(* IEC 61131-3 sources: daoli-st-library/DL_Device (part 7) *)

(* ---- I_DL_BarcodeScanner.st ---- *)
(*==============================================================================
 * 组件名称 (Component)  : I_DL_BarcodeScanner
 * 所属子库 (Sublibrary) : DL_Device
 * 当前版本 (Version)    : 1.0.0
 * 兼容性   (Platform)   : CODESYS 3.5 / TwinCAT 3 / 汇川 InoProShop / Machine Expert
 *                         纯 IEC 61131-3（第3版）接口语法，零厂商方言
 * 分类     (Category)   : 设备抽象接口（Interface）+ 配套状态枚举（DUT）
 * 功能简述 (Function)   : 工业固定式扫码枪标准抽象契约。路由分拣、批次追
 *                         溯、上下料校验等 DL_Process 模板的依赖注入件。
 *                         定义状态读取属性组（GET）与触发/应答/复位方法组；
 *                         串口/总线收发与数据本体由实现块（如
 *                         FB_DL_SerialScanner）经 IN_OUT 引脚注入，接口层
 *                         不做任何串口/总线收发与过程映像读写。
 * 契约结构 (Structure)  : 公约 0.11 接口三段式——状态枚举（本文件承载）+
 *                         属性（PROPERTY GET）+ 方法（METHOD）；方法共 3 个
 *                         （≤6 红线内）。故障态一律拒绝方法（红线：接口方
 *                         法拒绝语义），返回 FALSE 不静默成功。
 * 开源溯源 (Origin)     : 来源标签 tcopen-component / scanner-handshake
 *                         （RAW_NOTES_R7 S-2/S-3：TcOpen 组件接口分层思想
 *                         ——属性/方法分离契约与命令-应答握手语义，Apache
 *                         -2.0 公开资料，仅借鉴分层思想；接口命名、枚举编
 *                         号、方法签名 100% 本库独立设计，clean-room 未复
 *                         制源码）。
 * 归属说明 (Ownership)  : 本文件同时承载 E_DL_ScannerState 枚举定义，该枚
 *                         归属接口 I_DL_BarcodeScanner，与其同文件发布
 *                         （公约 0.11；禁止异文件同名异型重复定义）。
 * 红线自检 (Redline)    : R1 零全局变量表/外部变量引用 ✓｜R2 零物理 IO 地址 ✓
 *                         R3 纯 IEC 61131-3 ✓｜R4 N/A（契约件无运算）
 *                         R5 全成员中英双语同行注释 ✓｜R6 N/A（接口无状态机）
 *                         R7 N/A（无实例调用）｜R18 INTERFACE/END_INTERFACE
 *                         成对终结 ✓
 * 修订历史 (Revision)   :
 *   2026-11-15  v1.0.0  首版入库（Round 07 · DL_Device 扫码枪族接口件）
 *============================================================================*)

(*-----------------------------------------------------------------------------
 * 枚举: E_DL_ScannerState（归属接口 I_DL_BarcodeScanner，与其同文件）
 * 含义: 扫码枪握手状态机离散状态。编号步长 10 留空位便于后续插态而不破坏
 *       已有工程；eFault 取 99 保证排序末位（全库枚举编号惯例）。
 *----------------------------------------------------------------------------*)
TYPE E_DL_ScannerState :
(
    eIdle      := 0,    // 空闲待机：可受理解码触发 / Idle, ready to accept a decode trigger
    eTriggered := 10,   // 已触发：触发单拍输出已发出，等待下一拍进入读码 / Triggered, one-shot trigger output emitted
    eReading   := 20,   // 读码等待：结果窗口期内等待扫码枪回数 / Reading, waiting for the scanner reply inside the result window
    eOk        := 30,   // 解码成功：条码已锁存，等待应答消费 / Read OK, barcode latched, awaiting acknowledge
    eNoRead    := 40,   // 未读到：重试耗尽后的 NoRead 结果保持态 / NoRead, result hold state after retries exhausted
    eFault     := 99    // 故障锁存：连续 NoRead 超限/非法状态等，复位可尝试恢复 / Latched fault, reset may recover
) UINT;
END_TYPE

(*-----------------------------------------------------------------------------
 * 接口: I_DL_BarcodeScanner
 * 边界防错: 故障态一律拒绝方法；接口层不做任何串口/总线收发（数据本体经
 *           实现块 IN_OUT 引脚注入）；实现块负责握手编排与结果校验。
 *----------------------------------------------------------------------------*)
INTERFACE I_DL_BarcodeScanner

// ---- 属性段（全部只读 GET，实现块一一落地）----------------------------------

PROPERTY eState    : E_DL_ScannerState // 当前握手状态（Current handshake state），枚举见 E_DL_ScannerState
PROPERTY bReady    : BOOL              // 就绪可触发（Scanner ready），TRUE=处于可受理触发的状态 / TRUE = trigger acceptable
PROPERTY bReadOk   : BOOL              // 解码成功且结果有效（Read OK），TRUE=sBarcode 有效待消费 / TRUE = barcode valid and pending
PROPERTY bNoRead   : BOOL              // 未读到（NoRead），TRUE=重试耗尽未获得有效条码 / TRUE = no valid barcode after retries
PROPERTY sBarcode  : STRING(255)       // 最近有效条码字符串（Last valid barcode），长度 ≤255，bReadOk=TRUE 时有效 / Last valid barcode, valid when bReadOk
PROPERTY nReadCount: UDINT             // 累计成功解码次数（Total successful reads），复位不清零（追溯口径）/ Cumulative reads, preserved over reset
PROPERTY bFault    : BOOL              // 故障锁存中（Fault latched），显式排除信息级码（R21）/ TRUE = latched fault, info codes excluded
PROPERTY uErrorId  : UDINT             // 末次故障码（Last error code），0=无故障，段位 16#0003_xxxx / Last error code, family 16#0003_xxxx

// ---- 方法段（单发指令，返回受理/合法性结果）----------------------------------

METHOD CmdTrigger : BOOL // 触发一次解码（Trigger one decode），仅空闲态受理；非空闲/故障态拒绝返回 FALSE / Trigger one decode, accepted only in idle, rejected otherwise
VAR_INPUT
END_VAR

    END_METHOD

METHOD CmdAck : BOOL // 应答清除结果保持位（Acknowledge clears the result hold），eOk/eNoRead 态受理，为下一次解码前提 / Ack accepted in eOk/eNoRead
VAR_INPUT
END_VAR

    END_METHOD

METHOD CmdReset : BOOL // 复位故障（Reset fault），仅故障态受理返回 TRUE / Reset accepted only in fault state
VAR_INPUT
END_VAR

    END_METHOD
END_INTERFACE

(* ---- I_DL_Cylinder.st ---- *)
(*==============================================================================
 * 组件名称 (Component)  : I_DL_Cylinder
 * 所属子库 (Sublibrary) : DL_Device
 * 当前版本 (Version)    : 1.0.0
 * 兼容性   (Platform)   : CODESYS 3.5 / TwinCAT 3 / 汇川 InoProShop / Machine Expert
 *                         纯 IEC 61131-3（第3版）接口语法，零厂商方言
 * 分类     (Category)   : 设备抽象接口（Interface）+ 配套状态枚举（DUT）
 * 功能简述 (Function)   : 双电控气缸标准抽象契约。定义状态读取属性组（GET）与
 *                         动作指令方法组（Extend/Retract/Stop/Reset），供
 *                         DL_Process 全部机站动作层做依赖注入与解耦调用；
 *                         具体电磁阀输出与传感器采集由实现块（如
 *                         FB_DL_PneumaticCylinder）完成，接口层不做任何
 *                         过程映像读写，仅承载纯软件契约。
 * 开源溯源 (Origin)     : 来源标签 lbp-device（RAW_NOTES_R5 S-4：工业气动气缸
 *                         FB 设计指南 / LOGO! 气缸应用帖 / 双线圈互锁惯例，
 *                         公开教学文章，仅借鉴状态集合与故障分类等通用工程
 *                         语义；接口命名、方法签名按本库红线独立设计，
 *                         clean-room 未复制任何源码行）。
 * 红线自检 (Redline)    : R1 零全局变量表/外部变量引用 ✓｜R2 零物理 IO 地址 ✓
 *                         R3 纯 IEC 61131-3 ✓｜R5 全成员中英双语同行注释 ✓
 *                         R18 接口以 END_INTERFACE 成对终结 ✓
 * 归属说明 (Ownership)  : 本文件同时承载 E_DL_CylinderState 枚举定义，
 *                         该枚举归属接口 I_DL_Cylinder，与其同文件发布。
 * 修订历史 (Revision)   :
 *   2026-11-15  v1.0.0  首版入库（R5 轮 · DL_Device 开库）
 *============================================================================*)

(*-----------------------------------------------------------------------------
 * 枚举: E_DL_CylinderState（归属接口 I_DL_Cylinder，与其同文件）
 * 含义: 双电控气缸状态机离散状态。数值步长 10 留空位，便于后续插态
 *       而不破坏已有工程的持久化数值；eFault 取 99 保证排序末位。
 *----------------------------------------------------------------------------*)
TYPE E_DL_CylinderState :
(
    eIdle       := 0,    // 空闲稳态：双线圈全断，气缸保持当前位置 / Idle steady state, both coils off, cylinder holds position
    eExtending  := 10,   // 伸出动作中：伸出线圈得电，等待伸出到位反馈 / Extending, extend coil energized, waiting for extended feedback
    eExtended   := 20,   // 已伸出到位：伸出到位磁开确认的稳定终态 / Fully extended, confirmed by extended reed switch
    eRetracting := 30,   // 缩回动作中：缩回线圈得电，等待缩回到位反馈 / Retracting, retract coil energized, waiting for retracted feedback
    eRetracted  := 40,   // 已缩回到位：缩回到位磁开确认的稳定终态 / Fully retracted, confirmed by retracted reed switch
    eFault      := 99    // 故障锁存态：超时/传感器冲突/非法状态，仅复位可清 / Latched fault state, cleared only by reset
) UINT;
END_TYPE

(*-----------------------------------------------------------------------------
 * 接口: I_DL_Cylinder
 * 契约结构: 属性（PROPERTY GET）+ 方法（METHOD）两段式；方法总数 4 个，
 *           满足接口方法 ≤6 的拆分红线。所有方法均为非阻塞单发语义，
 *           不含跨扫描周期状态驻留；返回值仅表示"指令是否被受理"，
 *           实际动作完成以属性 eState/bExtended/bRetracted 为准。
 * 边界防错: 任何动作方法在故障锁存态一律拒绝并返回 FALSE；实现块负责
 *           信号采集与线圈驱动的全部过程映像交互，本接口不涉及。
 *----------------------------------------------------------------------------*)
INTERFACE I_DL_Cylinder

// ---- 属性段（全部只读 GET）------------------------------------------------

PROPERTY eState     : E_DL_CylinderState // 当前状态机状态（Current state）
PROPERTY bExtended  : BOOL               // 伸出到位磁开反馈（Extended reed feedback），TRUE=伸出到位
PROPERTY bRetracted : BOOL               // 缩回到位磁开反馈（Retracted reed feedback），TRUE=缩回到位
PROPERTY bFault     : BOOL               // 故障锁存中（Fault latched），TRUE=存在未复位故障
PROPERTY uErrorId   : UDINT              // 末次故障码（Last error code），0=无故障，段位 16#0003_xxxx

// ---- 方法段（单发指令，返回受理结果）--------------------------------------

METHOD CmdExtend : BOOL // 伸出指令（Extend command），单发；故障态拒绝返回 FALSE
VAR_INPUT
END_VAR

    END_METHOD

METHOD CmdRetract : BOOL // 缩回指令（Retract command），单发；故障态拒绝返回 FALSE
VAR_INPUT
END_VAR

    END_METHOD

METHOD CmdStop : BOOL // 停止指令（Stop command）：双线圈全断、保持当前位置；故障态拒绝返回 FALSE
VAR_INPUT
END_VAR

    END_METHOD

METHOD CmdReset : BOOL // 复位指令（Reset command），返回是否可复位（存在故障时为 TRUE）
VAR_INPUT
END_VAR

    END_METHOD
END_INTERFACE

(* ---- I_DL_FlowMeter.st ---- *)
(*==============================================================================
 * 组件名称 (Component)  : I_DL_FlowMeter
 * 所属子库 (Sublibrary) : DL_Device
 * 当前版本 (Version)    : 1.0.1
 * 兼容性   (Platform)   : CODESYS 3.5 / TwinCAT 3 / 汇川 InoProShop / Machine Expert
 *                         纯 IEC 61131-3（第3版）接口语法，零厂商方言
 * 分类     (Category)   : 设备抽象接口（Interface）+ 配套状态枚举（DUT）
 * 功能简述 (Function)   : 流量计标准抽象契约（脉冲型/模拟型均可适配）。定义
 *                         瞬时流量/累计总量读取属性组（GET）与总量清零/预置/
 *                         复位方法组，供批控与计量工站做依赖注入；脉冲采集
 *                         与频率估计由实现块（如 FB_DL_PulseFlowMeter）完成，
 *                         接口层不读物理输入。
 * 契约结构 (Structure)  : 公约 0.11 接口三段式——状态枚举（本文件承载）+
 *                         属性（PROPERTY GET）+ 方法（METHOD）；方法共 3 个
 *                         （≤6 红线内）。故障态一律拒绝方法。
 * 开源溯源 (Origin)     : 来源标签 tcopen-component / flow-totalizer
 *                         （RAW_NOTES_R7 S-2/S-6：TcOpen 组件接口分层思想与
 *                         工业流量计量公开语义域——瞬时流量/累计总量/低流
 *                         量截止，公开资料，仅借鉴语义域；接口命名、枚举编
 *                         号、方法签名 100% 本库独立设计，clean-room 未复
 *                         制源码）。
 * 归属说明 (Ownership)  : 本文件同时承载 E_DL_FlowMeterState 枚举定义，该枚
 *                         举归属接口 I_DL_FlowMeter，与其同文件发布（公约
 *                         0.11；禁止异文件同名异型重复定义）。
 * 红线自检 (Redline)    : R1 零全局变量表/外部变量引用 ✓｜R2 零物理 IO 地址 ✓
 *                         R3 纯 IEC 61131-3 ✓｜R4 N/A（契约件无运算）
 *                         R5 全成员中英双语同行注释 ✓｜R6 N/A（接口无状态机）
 *                         R7 N/A（无实例调用）｜R18 INTERFACE/END_INTERFACE
 *                         成对终结 ✓
 * 修订历史 (Revision)   :
 *   2026-11-15  v1.0.0  首版入库（Round 07 · DL_Device 流量计族接口件）
 *   2026-11-15  v1.0.1  R11 修复：枚举成员分隔符笔误，eFlowOk / eLowCutoff 两行误写单冒号 `:`（枚举成员赋值须用 `:=`），三平台编译阻断已消除，数值与语义不变。
 *                       R11 fix: enum member separator erratum, `:` -> `:=` on two members.
 *============================================================================*)

(*-----------------------------------------------------------------------------
 * 枚举: E_DL_FlowMeterState（归属接口 I_DL_FlowMeter，与其同文件）
 * 含义: 流量计量离散状态。编号步长 10 留空位，eFault 取 99 保证排序末位
 *       （全库枚举编号惯例）。
 *----------------------------------------------------------------------------*)
TYPE E_DL_FlowMeterState :
(
    eIdle      := 0,   // 空闲：未建窗或脉冲丢失超时后的静默态 / Idle, no window yet or silent after pulse timeout
    eMeasuring := 10,   // 测量中：采样窗运行中，流量待有效判定 / Measuring, sample window running, flow pending validation
    eFlowOk    := 20,  // 流量正常：高于低流量截止阈值的有效流量 / Flow OK, flow above the low-flow cutoff
    eLowCutoff := 30,  // 低流量截止：有效但低于阈值被截零（信息级）/ Low-flow cutoff, valid but zeroed below threshold (info)
    eFault     := 99   // 故障锁存：K 系数非法/非法状态，复位可尝试恢复 / Latched fault, reset may recover
) UINT;
END_TYPE

(*-----------------------------------------------------------------------------
 * 接口: I_DL_FlowMeter
 * 边界防错: 故障态一律拒绝方法并返回 FALSE；接口层不读物理输入；累计溢出
 *           防护（LREAL 整数精度边界预警）在实现块承载。
 *----------------------------------------------------------------------------*)
INTERFACE I_DL_FlowMeter

// ---- 属性段（全部只读 GET，实现块一一落地）----------------------------------

PROPERTY eState     : E_DL_FlowMeterState // 当前计量状态（Current metering state），枚举见 E_DL_FlowMeterState
PROPERTY fFlowRate  : REAL                // 瞬时流量（Flow rate）[L/min]，按 K 系数域换算 / Instantaneous flow rate [L/min], K-factor domain
PROPERTY fTotal     : LREAL               // 累计总量（Totalized volume）[L]，LREAL 防累计精度丢失 / Totalized volume [L], LREAL against precision loss
PROPERTY nPulseCount: UDINT               // 窗口内脉冲计数原始值（Pulse count of last window）/ Raw pulse count of the last window
PROPERTY bFault     : BOOL                // 故障锁存中（Fault latched），显式排除信息级码（R21）/ TRUE = latched fault, info codes excluded
PROPERTY uErrorId   : UDINT               // 末次故障码（Last error code），0=无故障，段位 16#0003_xxxx / Last error code, family 16#0003_xxxx

// ---- 方法段（单发指令，返回受理/合法性结果）----------------------------------

METHOD CmdTotalReset : BOOL // 总量清零（Total reset），批控切换零点；故障态拒绝 / Total reset, rejected in fault
VAR_INPUT
END_VAR

    END_METHOD

METHOD CmdTotalPreset : BOOL // 总量预置（Total preset），非有限值/负值拒绝 / Total preset, non-finite or negative rejected
VAR_INPUT
    fPreset : LREAL; // 预置总量（Preset volume）[L]，域 ≥0 / Preset volume [L], range >= 0
END_VAR

    END_METHOD

METHOD CmdReset : BOOL // 复位故障（Reset fault），仅故障态受理 / Reset accepted only in fault state
VAR_INPUT
END_VAR

    END_METHOD
END_INTERFACE

(* ---- I_DL_LevelSwitch.st ---- *)
(*==============================================================================
 * 组件名称 (Component)  : I_DL_LevelSwitch
 * 所属子库 (Sublibrary) : DL_Device
 * 当前版本 (Version)    : 1.0.0
 * 兼容性   (Platform)   : CODESYS 3.5 / TwinCAT 3 / 汇川 InoProShop / Machine Expert
 *                         纯 IEC 61131-3（第3版）接口语法，零厂商方言
 * 分类     (Category)   : 设备抽象接口（Interface）+ 配套状态枚举（DUT）
 * 功能简述 (Function)   : 料位开关标准抽象契约（振动叉/阻旋/电容等点式料位
 *                         开关通用）。高点溢流与低点干转联锁的统一契约；定
 *                         义有料判定/高/低联锁输出属性组（GET）与复位/测试
 *                         方法组；检测本体在传感器内部，接口层不做检测算法。
 * 契约结构 (Structure)  : 公约 0.11 接口三段式——状态枚举 + 失效安全模式枚
 *                         举（均本文件承载）+ 属性（PROPERTY GET）+ 方法
 *                         （METHOD）；方法共 2 个（≤6 红线内）。
 * 开源溯源 (Origin)     : 来源标签 tcopen-component / level-switch-failsafe
 *                         （RAW_NOTES_R7 S-2/S-7：TcOpen 组件接口分层思想与
 *                         料位开关失效安全公开语义域——fail-safe HIGH/LOW
 *                         方向约定、双联锁输出，公开资料，仅借鉴语义域；接
 *                         口命名、枚举编号、方法签名 100% 本库独立设计，
 *                         clean-room 未复制源码）。
 * 归属说明 (Ownership)  : 本文件同时承载 E_DL_LevelState 与 E_DL_FailSafeMode
 *                         两个枚举定义，均归属接口 I_DL_LevelSwitch，与其同
 *                         文件发布（公约 0.11；禁止异文件同名异型重复定义）。
 * 红线自检 (Redline)    : R1 零全局变量表/外部变量引用 ✓｜R2 零物理 IO 地址 ✓
 *                         R3 纯 IEC 61131-3 ✓｜R4 N/A（契约件无运算）
 *                         R5 全成员中英双语同行注释 ✓｜R6 N/A（接口无状态机）
 *                         R7 N/A（无实例调用）｜R18 INTERFACE/END_INTERFACE
 *                         成对终结 ✓
 * 修订历史 (Revision)   :
 *   2026-11-15  v1.0.0  首版入库（Round 07 · DL_Device 料位开关族接口件）
 *============================================================================*)

(*-----------------------------------------------------------------------------
 * 枚举: E_DL_LevelState（归属接口 I_DL_LevelSwitch，与其同文件）
 * 含义: 料位开关诊断状态。编号步长 10 留空位，eFault 取 99 保证排序末位
 *       （全库枚举编号惯例）。
 *----------------------------------------------------------------------------*)
TYPE E_DL_LevelState :
(
    eNoMaterial := 0,   // 无料：裸露确认态 / No material, bare confirmed
    eMaterial   := 10,  // 有料：覆盖确认态 / Material present, covered confirmed
    eSensorLoss := 20,  // 传感器失效态：按失效安全方向归一后的诊断镜像（本轮预留，检测算法后续轮次落地）/ Sensor loss, fail-safe normalized mirror (reserved this round)
    eFault      := 99   // 故障锁存：模式枚举越界等 / Latched fault
) UINT;
END_TYPE

(*-----------------------------------------------------------------------------
 * 枚举: E_DL_FailSafeMode（归属接口 I_DL_LevelSwitch，与其同文件）
 * 含义: 失效安全方向模式。决定传感器失效/使能切断时输出强制镜像的安全侧：
 *       eHigh=失效报有料（防溢流）；eLow=失效报无料（防干转）。
 *----------------------------------------------------------------------------*)
TYPE E_DL_FailSafeMode :
(
    eHigh := 0,   // 失效安全 HIGH：失效报有料，防溢流方向 / Fail-safe HIGH: failure reads covered, overflow protection
    eLow  := 1    // 失效安全 LOW：失效报无料，防干转方向 / Fail-safe LOW: failure reads bare, dry-run protection
) UINT;
END_TYPE

(*-----------------------------------------------------------------------------
 * 接口: I_DL_LevelSwitch
 * 边界防错: 故障态一律拒绝方法并返回 FALSE；接口层不做检测算法（检测本体
 *           在传感器内部）。
 *----------------------------------------------------------------------------*)
INTERFACE I_DL_LevelSwitch

// ---- 属性段（全部只读 GET，实现块一一落地）----------------------------------

PROPERTY eState    : E_DL_LevelState // 当前诊断状态（Current diagnostic state），枚举见 E_DL_LevelState
PROPERTY bMaterial : BOOL            // 有料判定输出（Material present），已按失效安全方向归一，TRUE=有料 / Fail-safe normalized material, TRUE = covered
PROPERTY bHighAlarm: BOOL            // 高点溢流联锁输出（High-level interlock），fail-safe HIGH 语义：归一有料即报警 / High alarm, fail-safe HIGH semantics
PROPERTY bLowAlarm : BOOL            // 低点干转联锁输出（Low-level interlock），fail-safe LOW 语义：归一无料即报警 / Low alarm, fail-safe LOW semantics
PROPERTY bFault    : BOOL            // 故障锁存中（Fault latched），显式排除信息级码（R21）/ TRUE = latched fault, info codes excluded
PROPERTY uErrorId  : UDINT           // 末次故障码（Last error code），0=无故障，段位 16#0003_xxxx / Last error code, family 16#0003_xxxx

// ---- 方法段（单发指令，返回受理/合法性结果）----------------------------------

METHOD CmdReset : BOOL // 复位故障（Reset fault），仅故障态受理 / Reset accepted only in fault state
VAR_INPUT
END_VAR

    END_METHOD

METHOD CmdTest : BOOL // 传感器功能测试请求（Sensor function test request），输出镜像进入测试态一拍 / Test request, test mirror asserted one scan
VAR_INPUT
END_VAR

    END_METHOD
END_INTERFACE

(* ---- I_DL_LightCurtain.st ---- *)
(*==============================================================================
 * 组件名称 (Component)  : I_DL_LightCurtain
 * 所属子库 (Sublibrary) : DL_Device
 * 当前版本 (Version)    : 1.0.0
 * 兼容性   (Platform)   : CODESYS 3.5 / TwinCAT 3 / 汇川 InoProShop / Machine Expert
 *                         纯 IEC 61131-3（第3版）接口语法，零厂商方言
 * 分类     (Category)   : 设备抽象接口（Interface）+ 配套状态枚举（DUT）
 * 功能简述 (Function)   : 安全光幕监控与屏蔽（Muting）标准抽象契约。定义光
 *                         幕状态读取属性组（GET）与滞留清除/确认/复位方法
 *                         组，供上层工站做依赖注入；OSSD 采集与屏蔽传感器
 *                         接线由实现块（如 FB_DL_SafetyLightCurtain）完成，
 *                         接口层不读物理输入。
 * 定位声明 (Positioning): 公约 0.13——本接口及其实现块为标准 PLC 逻辑编排
 *                         与诊断镜像层，不构成 ISO 13849 / IEC 62061 认证
 *                         安全功能，安全回路由认证安全控制器/安全 PLC 承载；
 *                         光幕本体 OSSD 的安全判断在认证安全光幕内部完成。
 * 契约结构 (Structure)  : 公约 0.11 接口三段式——状态枚举（本文件承载）+
 *                         属性（PROPERTY GET）+ 方法（METHOD）；方法共 3 个
 *                         （≤6 红线内）。故障态一律拒绝方法。
 * 边界防错 (Guard)      : bSafeStop 输出永不因屏蔽/override 置假——屏蔽态下
 *                         bSafeStop 断言恒 FALSE（光幕正常），实现块出口断
 *                         言承载。
 * 开源溯源 (Origin)     : 来源标签 tcopen-component / light-curtain-muting
 *                         （RAW_NOTES_R7 S-2/S-5：TcOpen 组件接口分层思想与
 *                         安全光幕屏蔽公开语义——OSSD 镜像、Muting/Override
 *                         状态域，公开资料，仅借鉴状态域语义；接口命名、枚
 *                         举编号、方法签名 100% 本库独立设计，clean-room 未
 *                         复制源码）。
 * 归属说明 (Ownership)  : 本文件同时承载 E_DL_CurtainState 枚举定义，该枚举
 *                         归属接口 I_DL_LightCurtain，与其同文件发布（公约
 *                         0.11；禁止异文件同名异型重复定义）。
 * 红线自检 (Redline)    : R1 零全局变量表/外部变量引用 ✓｜R2 零物理 IO 地址 ✓
 *                         R3 纯 IEC 61131-3 ✓｜R4 N/A（契约件无运算）
 *                         R5 全成员中英双语同行注释 ✓｜R6 N/A（接口无状态机）
 *                         R7 N/A（无实例调用）｜R18 INTERFACE/END_INTERFACE
 *                         成对终结 ✓
 * 修订历史 (Revision)   :
 *   2026-11-15  v1.0.0  首版入库（Round 07 · DL_Device 光幕族接口件）
 *============================================================================*)

(*-----------------------------------------------------------------------------
 * 枚举: E_DL_CurtainState（归属接口 I_DL_LightCurtain，与其同文件）
 * 含义: 光幕监控/屏蔽离散状态。编号步长 10 留空位，eFault 取 99 保证排序末
 *       位（全库枚举编号惯例）。
 *----------------------------------------------------------------------------*)
TYPE E_DL_CurtainState :
(
    eClear    := 0,   // 通光：光幕未被遮挡且无屏蔽活动 / Clear, curtain unblocked and no muting activity
    eBlocked  := 10,  // 遮挡：光幕被遮挡且未屏蔽（应停机镜像态）/ Blocked, curtain interrupted without muting (safe-stop mirror)
    eMuting   := 20,  // 屏蔽进行中：合法屏蔽序列屏蔽中 / Muting, a legal muting sequence is active
    eOverride := 30,   // 滞留清除进行中：钥匙开关滞留物清除 / Override, key-switch residual-object clearing active
    eFault    := 99   // 故障锁存：序列错误/屏蔽超时/OSSD 不一致/非法状态 / Latched fault
) UINT;
END_TYPE

(*-----------------------------------------------------------------------------
 * 接口: I_DL_LightCurtain
 * 边界防错: 故障态一律拒绝方法并返回 FALSE；bSafeStop 永不因屏蔽/override
 *           置假（屏蔽态下断言恒 FALSE，实现块承载）。
 *----------------------------------------------------------------------------*)
INTERFACE I_DL_LightCurtain

// ---- 属性段（全部只读 GET，实现块一一落地）----------------------------------

PROPERTY eState         : E_DL_CurtainState // 当前光幕状态（Current curtain state），枚举见 E_DL_CurtainState
PROPERTY bClear         : BOOL              // 光幕通光（Clear），OSSD 双通道全通光 / OSSD both channels clear
PROPERTY bMutingActive  : BOOL              // 屏蔽进行中（Muting active），合法屏蔽序列屏蔽中 / TRUE = legal muting sequence active
PROPERTY bOverrideActive: BOOL              // 滞留清除进行中（Override active），滞留物清除中 / TRUE = override clearing active
PROPERTY bSafeStop      : BOOL              // 应停机输出（Safe stop），光幕被遮挡且未屏蔽——本接口核心安全镜像位 / Curtain blocked and not muted, core safe-stop mirror
PROPERTY bFault         : BOOL              // 故障锁存中（Fault latched），显式排除信息级码（R21）/ TRUE = latched fault, info codes excluded
PROPERTY uErrorId       : UDINT             // 末次故障码（Last error code），0=无故障，段位 16#0003_xxxx / Last error code, family 16#0003_xxxx

// ---- 方法段（单发指令，返回受理/合法性结果）----------------------------------

METHOD CmdOverride : BOOL // 滞留物清除请求（Override request），前提至少一个屏蔽传感器仍遮挡，否则拒绝 / Override accepted only with at least one muting sensor blocked
VAR_INPUT
END_VAR

    END_METHOD

METHOD CmdAck : BOOL // 屏蔽/故障确认复位（Acknowledge of muting abort/fault），屏蔽序列中止后回评估态受理 / Ack after a muting abort, back to evaluation
VAR_INPUT
END_VAR

    END_METHOD

METHOD CmdReset : BOOL // 复位故障与重启联锁（Reset fault and restart interlock），仅故障态受理 / Reset accepted only in fault state
VAR_INPUT
END_VAR

    END_METHOD
END_INTERFACE

(* ---- I_DL_MotorDriver.st ---- *)
(*==============================================================================
 * 组件名称 (Component)  : I_DL_MotorDriver
 * 所属子库 (Sublibrary) : DL_Device
 * 当前版本 (Version)    : 1.0.0
 * 兼容性   (Platform)   : CODESYS 3.5 / TwinCAT 3 / 汇川 InoProShop / Machine Expert
 *                         纯 IEC 61131-3（第3版）接口语法，零厂商方言
 * 分类     (Category)   : 设备抽象接口（Interface）+ 配套状态枚举（DUT）
 * 功能简述 (Function)   : 直接启动（DOL）电机驱动器标准抽象契约。定义状态
 *                         读取属性组（GET，含重启抑制指示）与启停/复位方法组，
 *                         供机站动作层与配电监控层做依赖注入与解耦调用；
 *                         接触器线圈驱动与反馈采集由实现块（如 FB_DL_DolMotor）
 *                         完成，接口层不做任何过程映像读写。
 * 开源溯源 (Origin)     : 来源标签 lbp-device（RAW_NOTES_R5 S-4：DOL 电机保护
 *                         惯例——接触器反馈校验窗、热继电器过载锁存、防频繁
 *                         启停与重启抑制冷却时间为行业公知语义，公开教学
 *                         资料，仅借鉴通用工程语义；接口命名、方法签名按
 *                         本库红线独立设计，clean-room 未复制源码）。
 * 红线自检 (Redline)    : R1 零全局变量表/外部变量引用 ✓｜R2 零物理 IO 地址 ✓
 *                         R3 纯 IEC 61131-3 ✓｜R5 全成员中英双语同行注释 ✓
 *                         R18 接口以 END_INTERFACE 成对终结 ✓
 * 归属说明 (Ownership)  : 本文件同时承载 E_DL_MotorState 枚举定义，
 *                         该枚举归属接口 I_DL_MotorDriver，与其同文件发布。
 * 修订历史 (Revision)   :
 *   2026-11-15  v1.0.0  首版入库（R5 轮 · DL_Device 开库）
 *============================================================================*)

(*-----------------------------------------------------------------------------
 * 枚举: E_DL_MotorState（归属接口 I_DL_MotorDriver，与其同文件）
 * 含义: DOL 电机驱动状态机离散状态。数值步长 10 留空位，便于后续插态
 *       而不破坏已有工程的持久化数值；eFault 取 99 保证排序末位。
 *----------------------------------------------------------------------------*)
TYPE E_DL_MotorState :
(
    eIdle          := 0,    // 空闲停机态：接触器断开，可受理启动指令 / Idle stopped state, contactor open, start commands accepted
    eStarting      := 10,   // 启动校验态：线圈已得电，等待反馈窗内触点吸合确认 / Starting, coil energized, awaiting contactor pick-up confirmation within feedback window
    eRunning       := 20,   // 运行态：反馈吸合确认，正常带载运行 / Running, contactor feedback confirmed, loaded operation
    eStopping      := 30,   // 停机过渡态：线圈已断，等待反馈触点分断确认 / Stopping transition, coil de-energized, awaiting contactor drop-out confirmation
    eTripOverload  := 40,   // 过载脱扣态：热继电器动作锁存，仅复位且过载信号消失后可清 / Overload tripped and latched, cleared only by reset with overload signal removed
    eFault         := 99    // 故障锁存态：拒动/失反馈等故障，仅复位可清 / Latched fault state (refusal, feedback loss), cleared only by reset
) UINT;
END_TYPE

(*-----------------------------------------------------------------------------
 * 接口: I_DL_MotorDriver
 * 契约结构: 属性（PROPERTY GET）+ 方法（METHOD）两段式；方法总数 3 个，
 *           满足接口方法 ≤6 的拆分红线。所有方法均为非阻塞单发语义，
 *           不含跨扫描周期状态驻留；启动/复位方法返回值表示"指令是否
 *           被受理"，实际运行状态以属性 eState/bRunning 为准。
 * 边界防错: 启动方法在被抑制（重启抑制/次数超限）或故障态一律返回 FALSE；
 *           停止为无条件安全指令；实现块负责线圈驱动与触点反馈采集的
 *           全部过程映像交互，本接口不涉及。
 *----------------------------------------------------------------------------*)
INTERFACE I_DL_MotorDriver

// ---- 属性段（全部只读 GET）------------------------------------------------

PROPERTY eState          : E_DL_MotorState // 当前状态机状态（Current state）
PROPERTY bRunning        : BOOL            // 运行反馈（Running feedback），TRUE=反馈吸合确认运行中 / TRUE = running confirmed by contactor feedback
PROPERTY bFault          : BOOL            // 故障锁存中（Fault latched），TRUE=存在未复位故障（含过载脱扣）/ TRUE = latched fault incl. overload trip
PROPERTY uErrorId        : UDINT           // 末次故障码（Last error code），0=无故障，段位 16#0003_xxxx / Last error code, 0 = none, family 16#0003_xxxx
PROPERTY bRestartInhibit : BOOL            // 重启抑制激活中（Restart inhibit active），TRUE=冷却期内拒绝启动 / TRUE = start refused during cooling period

// ---- 方法段（单发指令，返回受理结果）--------------------------------------

METHOD CmdStart : BOOL // 启动指令（Start command），单发；被抑制/故障态返回 FALSE / Rejected with FALSE when inhibited or faulty
VAR_INPUT
END_VAR

    END_METHOD

METHOD CmdStop // 停止指令（Stop command），无条件安全动作，双线圈全断 / Unconditional safe stop command
VAR_INPUT
END_VAR

    END_METHOD

METHOD CmdReset : BOOL // 复位过载/故障（Reset overload and fault），返回是否可复位 / Returns TRUE only when resettable
VAR_INPUT
END_VAR

    END_METHOD
END_INTERFACE

(* ---- I_DL_MotorizedValve.st ---- *)
(*==============================================================================
 * 组件名称 (Component)  : I_DL_MotorizedValve
 * 所属子库 (Sublibrary) : DL_Device
 * 当前版本 (Version)    : 1.0.0
 * 兼容性   (Platform)   : CODESYS 3.5 / TwinCAT 3 / 汇川 InoProShop / Machine Expert
 *                         纯 IEC 61131-3（第3版）接口语法，零厂商方言
 * 分类     (Category)   : 设备抽象接口（Interface）+ 配套状态枚举（DUT）
 * 功能简述 (Function)   : 电动调节阀（开/关脉冲输出、无阀位变送器）标准
 *                         抽象契约。定义状态读取属性组（GET）与开阀/关阀/
 *                         停止/复位方法组，供暖通水路与工艺管路的调节
 *                         回路做依赖注入与解耦调用；双脉冲输出、行程时间
 *                         积分估算与限位保护由实现块（如
 *                         FB_DL_ThreePointValve）完成，接口层不做任何
 *                         过程映像读写，仅承载纯软件契约。
 * 开源溯源 (Origin)     : 来源标签 lbp-basic-process / lbp-device
 *                         （RAW_NOTES_R6 S-1 + S-5：三点浮点式电动阀的开/
 *                         关脉冲控制惯例、行程时间开度估算语义等行业
 *                         公知工程惯例，公开教学资料，仅借鉴通用工程语义；
 *                         接口命名、方法签名按本库红线独立设计，clean-room
 *                         未复制源码）。
 * 红线自检 (Redline)    : R1 零全局变量表/外部变量引用 ✓｜R2 零物理 IO 地址 ✓
 *                         R3 纯 IEC 61131-3 ✓｜R5 全成员中英双语同行注释 ✓
 *                         R18 接口以 END_INTERFACE 成对终结 ✓
 * 归属说明 (Ownership)  : 本文件同时承载 E_DL_MotorValveState 枚举定义，
 *                         该枚举归属接口 I_DL_MotorizedValve，与其同文件
 *                         发布。
 * 修订历史 (Revision)   :
 *   2026-11-15  v1.0.0  首版入库（R6 轮 · DL_Device 阀门/驱动族深化）
 *============================================================================*)

(*-----------------------------------------------------------------------------
 * 枚举: E_DL_MotorValveState（归属接口 I_DL_MotorizedValve，与其同文件）
 * 含义: 电动调节阀状态机离散状态。数值步长 10 留空位，便于后续插态
 *       而不破坏已有工程的持久化数值；eFault 取 99 保证排序末位。
 *----------------------------------------------------------------------------*)
TYPE E_DL_MotorValveState :
(
    eIdle    := 0,    // 空闲稳态：双脉冲全断，阀停在当前位置 / Idle steady state, both pulses off, valve holds position
    eOpening := 10,   // 开阀中：开阀脉冲输出，行程时间积分估算开度 / Opening, open pulse active, position integrated from stroke time
    eClosing := 20,   // 关阀中：关阀脉冲输出，行程时间积分估算开度 / Closing, close pulse active, position integrated from stroke time
    eOpened  := 30,   // 全开确认：全开限位反馈确认的端点稳态 / Fully opened, endpoint confirmed by open limit switch
    eClosed  := 40,   // 全关确认：全关限位反馈确认的端点稳态 / Fully closed, endpoint confirmed by closed limit switch
    eFault   := 99    // 故障锁存态：估算失准/限位冲突/非法状态，仅复位可清 / Latched fault state, cleared only by reset
) UINT;
END_TYPE

(*-----------------------------------------------------------------------------
 * 接口: I_DL_MotorizedValve
 * 契约结构: 属性（PROPERTY GET）+ 方法（METHOD）两段式；方法总数 4 个，
 *           满足接口方法 ≤6 的拆分红线。所有方法均为非阻塞单发语义，
 *           不含跨扫描周期状态驻留；返回值仅表示"指令是否被受理"，
 *           实际阀位以属性 eState/fPosEstimate 为准。
 * 边界防错: 故障态下动作方法一律拒绝并返回 FALSE；已在端点（限位确认）
 *           的指令受理但由实现块拒绝执行并置信息级；实现块负责双脉冲
 *           输出与限位采集的全部过程映像交互，本接口不涉及。
 *----------------------------------------------------------------------------*)
INTERFACE I_DL_MotorizedValve

// ---- 属性段（全部只读 GET）------------------------------------------------

PROPERTY eState       : E_DL_MotorValveState // 当前状态机状态（Current state）
PROPERTY fPosEstimate : REAL          // 估算开度（Estimated position）[%]，0~100，由行程时间积分自动估算 / Estimated position [%], integrated from stroke time
PROPERTY bLimOpen     : BOOL          // 全开限位反馈（Open limit switch），TRUE=已到全开端点 / TRUE = at fully-open endpoint
PROPERTY bLimClosed   : BOOL          // 全关限位反馈（Closed limit switch），TRUE=已到全关端点 / TRUE = at fully-closed endpoint
PROPERTY bFault       : BOOL          // 故障锁存中（Fault latched），TRUE=存在未复位故障 / TRUE = latched fault present
PROPERTY uErrorId     : UDINT         // 末次事件码（Last error code），0=无，段位 16#0003_xxxx / Last error code, 0 = none, family 16#0003_xxxx

// ---- 方法段（单发指令，返回受理结果）--------------------------------------

METHOD CmdOpen : BOOL // 开阀指令（Open command），电平语义受理为保持锁存；故障态拒绝返回 FALSE / Open command held as latch, rejected in fault
VAR_INPUT
END_VAR

    END_METHOD

METHOD CmdClose : BOOL // 关阀指令（Close command），电平语义受理为保持锁存；故障态拒绝返回 FALSE / Close command held as latch, rejected in fault
VAR_INPUT
END_VAR

    END_METHOD

METHOD CmdStop : BOOL // 双脉冲全断保持（Stop command, both pulses off, hold position）；无条件受理 / Unconditionally accepted
VAR_INPUT
END_VAR

    END_METHOD

METHOD CmdReset : BOOL // 复位指令（Reset command），返回是否可复位（存在故障时为 TRUE）/ Returns TRUE only when resettable
VAR_INPUT
END_VAR

    END_METHOD
END_INTERFACE

(* ---- I_DL_ProportionalValve.st ---- *)
(*==============================================================================
 * 组件名称 (Component)  : I_DL_ProportionalValve
 * 所属子库 (Sublibrary) : DL_Device
 * 当前版本 (Version)    : 1.0.0
 * 兼容性   (Platform)   : CODESYS 3.5 / TwinCAT 3 / 汇川 InoProShop / Machine Expert
 *                         纯 IEC 61131-3（第3版）接口语法，零厂商方言
 * 分类     (Category)   : 设备抽象接口（Interface）+ 配套状态枚举（DUT）
 * 功能简述 (Function)   : 模拟量比例阀/调节阀（开度指令-反馈型）标准抽象
 *                         契约。定义状态读取属性组（GET）与阀位设定/停止/
 *                         复位方法组，供温度、流量、压力等过程调节回路
 *                         做依赖注入与解耦调用；指令整形、限幅域映射与
 *                         反馈诊断由实现块（如 FB_DL_AnalogValve）完成，
 *                         接口层不做任何过程映像读写，仅承载纯软件契约。
 * 开源溯源 (Origin)     : 来源标签 lbp-basic-process / lbp-device
 *                         （RAW_NOTES_R6 S-1：比例调节阀开度指令-反馈控制
 *                         惯例、偏差报警语义等行业公知工程惯例，公开教学
 *                         资料，仅借鉴通用工程语义；接口命名、方法签名按
 *                         本库红线独立设计，clean-room 未复制源码）。
 * 红线自检 (Redline)    : R1 零全局变量表/外部变量引用 ✓｜R2 零物理 IO 地址 ✓
 *                         R3 纯 IEC 61131-3 ✓｜R5 全成员中英双语同行注释 ✓
 *                         R18 接口以 END_INTERFACE 成对终结 ✓
 * 归属说明 (Ownership)  : 本文件同时承载 E_DL_ValveState 枚举定义，该枚举
 *                         归属接口 I_DL_ProportionalValve，与其同文件发布。
 * 修订历史 (Revision)   :
 *   2026-11-15  v1.0.0  首版入库（R6 轮 · DL_Device 阀门/驱动族深化）
 *============================================================================*)

(*-----------------------------------------------------------------------------
 * 枚举: E_DL_ValveState（归属接口 I_DL_ProportionalValve，与其同文件）
 * 含义: 比例调节阀状态机离散状态。数值步长 10 留空位，便于后续插态
 *       而不破坏已有工程的持久化数值；eFault 取 99 保证排序末位。
 *----------------------------------------------------------------------------*)
TYPE E_DL_ValveState :
(
    eIdle        := 0,    // 空闲稳态：调节使能撤除或输出冻结，保持当前阀位 / Idle steady state, modulating disabled or output frozen, holds position
    eModulating  := 10,   // 调节中：调节使能有效，阀位指令整形后正常输出 / Modulating, enable active, position command shaping and output active
    eFault       := 99    // 故障锁存态：反馈失效/非法状态，仅复位可清 / Latched fault state (feedback loss), cleared only by reset
) UINT;
END_TYPE

(*-----------------------------------------------------------------------------
 * 接口: I_DL_ProportionalValve
 * 契约结构: 属性（PROPERTY GET）+ 方法（METHOD）两段式；方法总数 3 个，
 *           满足接口方法 ≤6 的拆分红线。所有方法均为非阻塞单发语义，
 *           不含跨扫描周期状态驻留；返回值仅表示"指令是否被受理/
 *           参数是否合法"，实际阀位以属性 fPosCmd/fPosFeedback 为准。
 * 边界防错: 设定方法在故障态拒绝并返回 FALSE；停止方法冻结输出保持
 *           当前阀位；实现块负责指令整形与反馈诊断的全部过程映像
 *           交互，本接口不涉及。
 *----------------------------------------------------------------------------*)
INTERFACE I_DL_ProportionalValve

// ---- 属性段（全部只读 GET）------------------------------------------------

PROPERTY eState          : E_DL_ValveState // 当前状态机状态（Current state）
PROPERTY fPosCmd         : REAL            // 当前阀位指令（Current position command）[%]，整形钳位后生效值 / Effective position command [%] after shaping
PROPERTY fPosFeedback    : REAL            // 阀位反馈（Position feedback）[%]，非有限值时保持末次有效值 / Position feedback [%], holds last valid on non-finite input
PROPERTY bDeviationAlarm : BOOL            // 偏差报警激活中（Deviation alarm），瞬时型每拍重算 / Transient deviation alarm, recomputed each cycle
PROPERTY bFault          : BOOL            // 故障锁存中（Fault latched），TRUE=存在未复位故障 / TRUE = latched fault present
PROPERTY uErrorId        : UDINT           // 末次事件码（Last error code），0=无，段位 16#0003_xxxx / Last error code, 0 = none, family 16#0003_xxxx

// ---- 方法段（单发指令，返回受理/合法性结果）--------------------------------

METHOD SetPosition : BOOL // 阀位指令设定（Position set）[%]，越界/非有限值拒绝并返回 FALSE / Position set command, out-of-range or non-finite returns FALSE
VAR_INPUT
    fPos : REAL; // 阀位设定值（Position value）[%]，域 0..100 / Position value [%], range 0..100
END_VAR

    END_METHOD

METHOD CmdStop : BOOL // 停止指令（Stop command）：冻结输出保持当前阀位，直至下次设定或使能撤除；故障态拒绝返回 FALSE / Freeze output until next set or enable drop, rejected in fault
VAR_INPUT
END_VAR

    END_METHOD

METHOD CmdReset : BOOL // 复位指令（Reset command），返回是否可复位（存在故障时为 TRUE）/ Returns TRUE only when resettable
VAR_INPUT
END_VAR

    END_METHOD
END_INTERFACE

(* ---- I_DL_RfidReader.st ---- *)
(*==============================================================================
 * 组件名称 (Component)  : I_DL_RfidReader
 * 所属子库 (Sublibrary) : DL_Device
 * 当前版本 (Version)    : 1.0.0
 * 组件分类 (Category)   : 接口（INTERFACE）+ 配套结构体与枚举（同文件发布）
 * 兼容性   (Platform)   : CODESYS 3.5 / TwinCAT 3 / 汇川 InoProShop / Schneider
 *                         Machine Expert；纯 IEC 61131-3 第 3 版接口语法，
 *                         零厂商方言，零标准库依赖
 * 功能描述 (Function)   : 载具与托盘 RFID 读写头的标准抽象契约。按本库接口
 *                         三段式组织（结构体 + 只读属性 + 单发方法），上层工站
 *                         只依赖本接口引用，即可用同一套代码适配串口读写头、
 *                         工业以太网读写头、IO-Link 读写头与仿真器。
 * 参数分段 (Segments)   : 借 AOI 的参数分段范式把接口切为四段：
 *                         In 段（指令）= 四个单发方法；
 *                         Out 段（状态）= 三个只读属性；
 *                         InOut 段（诊断与组态）= ST_DL_RfidDiag 与 ST_DL_RfidCfg
 *                         经属性与方法参数整体吞吐；
 *                         Local 段（内部中间量）= 留给实现块，接口不出现。
 *                         只借分段组织与访问等级思想，未接触任何厂商的 UDT
 *                         布局、参数命名与内部逻辑。
 * 与既有件边界 (Boundary): I_DL_BarcodeScanner 是一维码扫描（触发应答握手、
 *                         单向只读）；本接口是读写双向加载具数据区（分页与
 *                         字块）加防重复读，方法语义与数据模型都不同，
 *                         不做继承合并。
 * 方法数红线 (Budget)   : 方法 4 个（Init / ReadTag / WriteTag / Reset），
 *                         属性 3 个（State / Tag / Diag），属性不计入方法预算
 *                         （与 I_DL_MotionAxis 同一口径），故满足接口方法数
 *                         不超过 6 的红线。
 * 语义约定 (Semantics)  :
 *   1 未 Init 或 Init 失败时，除 Reset 与三个只读属性外全部方法返回 FALSE 并
 *     给出非零码，且不改变任何内部状态；
 *   2 全部方法为非阻塞单发：方法内只登记请求并置内部标志，跨周期动作由实现块
 *     主体状态机执行，方法内不得出现等待循环；
 *   3 忙态（内部指令执行中）再调用 ReadTag 或 WriteTag 一律返回 FALSE 并给码，
 *     不排队不缓存（读头硬件本身互斥，排队只会让上层误以为指令已生效）；
 *   4 视野内无标签是业务态不是故障：不置故障位、不进故障态、不计入重试次数；
 *   5 所有失败必须区分「组态或使用类」与「工艺类」两类码段，HMI 据此决定是
 *     叫工程师改参数还是叫维修换硬件。
 * 开源溯源 (Origin)     : tcopen-component / rockwell-aoi。参考 TcOpen 公开组件
 *                         库的契约与实现分离范式（接口只定义成员签名，状态经
 *                         只读属性暴露），以及 Rockwell AOI 公开手册所述的参数
 *                         分段与外部访问等级思想（Instruction / Status /
 *                         InOut / Local 四段，Input 与 Output 只读、InOut 与
 *                         Local 对外不可见）。仅借分段组织与访问等级，结构体
 *                         布局、成员命名、码位与状态机 100% 自有 clean-room，
 *                         不构成衍生作品。
 * 依赖     (Depends)    : 无 DL_ 内部依赖；无标准库功能块依赖
 * 归属声明 (Ownership)  : 本文件同时承载 E_DL_RfidState、ST_DL_RfidTag、
 *                         ST_DL_RfidDiag、ST_DL_RfidCfg 四个类型定义，均归属
 *                         本接口并与其同文件发布（库内公约 0.18）。
 * 修订历史 (Revision)   :
 *   2026-11-15  v1.0.0  首版入库（Round 10 · T2-6 Rockwell AOI 开组）
 *============================================================================*)

(*------------------------------------------------------------------------------
 * 枚举: E_DL_RfidState
 * 含义: 对外可观测的读写头状态。区间 0 到 20 为常规态，90 以上为异常与业务态，
 *       数值步长 10 留空位，新增状态不破坏已有 HMI 的数值映射
 *-----------------------------------------------------------------------------*)
TYPE E_DL_RfidState :
(
    eOffline := 0,     // 未初始化或未上电：除复位与只读属性外全部拒绝 / Offline, only reset and read-only members are served
    eReady   := 10,    // 就绪，可受理指令 / Ready, accepts commands
    eBusy    := 20,    // 指令执行中，互斥，禁止重入 / Busy, mutually exclusive, re-entry rejected
    eError   := 90,    // 故障，需复位清除 / Fault, cleared only by reset
    eNoTag   := 95     // 视野内无标签，业务态非故障 / No tag in field, a business state rather than a fault
);
END_TYPE

(*------------------------------------------------------------------------------
 * 结构体: ST_DL_RfidTag
 * 含义: 一次读写的标签快照。读到后保持（R27），直到下次成功读取覆盖
 *-----------------------------------------------------------------------------*)
TYPE ST_DL_RfidTag :
STRUCT
    sTagId  : STRING(64);   // 标签唯一号，空串表示无标签 [ASCII] / Tag unique identifier, empty means no tag
    sData   : STRING(64);   // 标签数据区内容，编码由组态决定 [ASCII 或十六进制] / Tag data area content
    uPage   : UINT;         // 数据页号，0 表示连续区 [页] / Data page number, zero means the contiguous area
    nRssi   : INT;          // 信号强度，域零下 90 到 0 [分贝毫瓦] / Signal strength, -90 to 0 dBm
    bValid  : BOOL;         // 本次读取有效 [-] / TRUE when this snapshot holds a valid read
END_STRUCT
END_TYPE

(*------------------------------------------------------------------------------
 * 结构体: ST_DL_RfidDiag
 * 含义: 诊断与统计。整体经只读属性回读，等价于 AOI 的 InOut 段对外封装
 *-----------------------------------------------------------------------------*)
TYPE ST_DL_RfidDiag :
STRUCT
    uLastErrorId : UDINT;   // 末次故障码，段位由实现块按子库公约自定 [代码] / Last error code, family defined by the implementer
    nCommRetry   : INT;     // 本次指令累计通信重试次数 [次] / Retry count of the current command
    nReadTotal   : DINT;    // 累计读成功次数，跨班不清零 [次] / Total successful reads, never cleared per shift
    nWriteTotal  : DINT;    // 累计写成功次数，跨班不清零 [次] / Total successful writes, never cleared per shift
    bAntennaOk   : BOOL;    // 天线自检通过 [-] / TRUE when the antenna self-test passed
    tLastComm    : TIME;    // 末次成功通信距今时长 [毫秒] / Elapsed time since the last successful communication
END_STRUCT
END_TYPE

(*------------------------------------------------------------------------------
 * 结构体: ST_DL_RfidCfg
 * 含义: 组态参数，调用方持有并经 Init 方法的 VAR_IN_OUT 注入，接口侧只读使用
 *-----------------------------------------------------------------------------*)
TYPE ST_DL_RfidCfg :
STRUCT
    sAntennaNo   : STRING(8);          // 天线号，多天线读头用于选天线 [ASCII] / Antenna selector for multi-antenna readers
    nPowerDbm    : INT;                // 发射功率，域 0 到 30 [分贝毫瓦] / Transmit power, 0 to 30 dBm
    tTimeout     : TIME;               // 单次指令超时，域 50 毫秒到 5 秒 [毫秒] / Per-command timeout, 50 ms to 5 s
    nMaxRetry    : INT;                // 重试次数，域 0 到 5 [次] / Retry count, 0 to 5
    bDupFilterEn : BOOL;               // 同标签重复读抑制使能 [-] / Duplicate-read suppression enable
    tDupWindow   : TIME;               // 重复读抑制窗，域 100 毫秒到 60 秒 [毫秒] / Duplicate suppression window
END_STRUCT
END_TYPE

(*------------------------------------------------------------------------------
 * 接口: I_DL_RfidReader
 * 契约结构: 属性段（只读 GET，Out 段）+ 方法段（单发，In 段）
 *-----------------------------------------------------------------------------*)
INTERFACE I_DL_RfidReader

// ---- 属性段（Out 段，全部只读，实现块以同名 PROPERTY GET 落地） -----------

PROPERTY State : E_DL_RfidState      // 当前状态，映射规则由实现块逐条写死（Current state, mapping fixed by the implementer）
PROPERTY Tag   : ST_DL_RfidTag       // 当前标签快照，读到后保持（Current tag snapshot, held after a successful read）
PROPERTY Diag  : ST_DL_RfidDiag      // 诊断结构整体回读（Whole diagnostic structure, read back at once）

// ---- 方法段（In 段，全部非阻塞单发，返回 FALSE 时必须给出非零码） --------

METHOD Init : BOOL                   // 初始化，组态经 VAR_IN_OUT 注入，只登记不阻塞（Initialise; configuration injected by reference）
VAR_IN_OUT
    stCfg : ST_DL_RfidCfg;           // 组态结构，调用方持有，接口侧只读 [结构] / Configuration structure owned by the caller, read-only here
END_VAR

    END_METHOD

METHOD ReadTag : BOOL                // 发起读标签（唯一号与数据区），忙时拒绝（Start a tag read, rejected while busy）
VAR_INPUT
END_VAR

    END_METHOD

METHOD WriteTag : BOOL               // 发起写数据区，内容经 VAR_IN_OUT 注入，忙时拒绝（Start a data write, rejected while busy）
VAR_IN_OUT
    stTagIn : ST_DL_RfidTag;         // 待写内容，实现块须锁存副本防调用方中途改动 [结构] / Payload to write; the implementer must latch a copy
END_VAR

    END_METHOD

METHOD Reset : BOOL                  // 清故障回就绪态，是故障态下唯一受理的方法（Clear the fault and return to ready）
VAR_INPUT
END_VAR

(*==============================================================================
 * 调用示例 (Instance guide)：
 *   VAR fbReader : FB_DL_RfidTagHandler;    // 具体实现块
 *       stCfg    : ST_DL_RfidCfg;           // 组态，调用方持有
 *       stTag    : ST_DL_RfidTag;           // 标签快照
 *       iReader  : I_DL_RfidReader;         // 接口引用，注入实现块
 *   END_VAR
 *   fbReader(stCfg := stCfg, bHwReady := bReaderReady);
 *   iReader := fbReader;                     // 依赖注入，上层只依赖接口
 *   IF iReader.State = E_DL_RfidState.eReady THEN
 *       bOk := iReader.ReadTag();
 *   END_IF
 *   IF iReader.Tag.bValid THEN
 *       sPalletId := iReader.Tag.sTagId;     // 保持型，读到后立即可用
 *   END_IF
 *   上层工站不得直接引用实现块类型，只能持有接口引用，替换硬件时只改注入点。
 *============================================================================*)

    END_METHOD
END_INTERFACE

(* ---- I_DL_SafetyDoor.st ---- *)
(*==============================================================================
 * 组件名称 (Component)  : I_DL_SafetyDoor
 * 所属子库 (Sublibrary) : DL_Device
 * 当前版本 (Version)    : 1.0.0
 * 兼容性   (Platform)   : CODESYS 3.5 / TwinCAT 3 / 汇川 InoProShop / Machine Expert
 *                         纯 IEC 61131-3（第3版）接口语法，零厂商方言
 * 分类     (Category)   : 设备抽象接口（Interface）+ 配套状态枚举（DUT）
 * 功能简述 (Function)   : 安全门联锁标准抽象契约（电磁锁扣门）。定义解锁时
 *                         序状态读取属性组（GET）与请求解锁/重新闭锁/复位/
 *                         审计清除方法组，供上层工站做依赖注入；电磁铁输出、
 *                         反馈采集与物理输出全部由实现块（如
 *                         FB_DL_GuardLockDoor）完成，接口层不写物理输出。
 * 定位声明 (Positioning): 公约 0.13——本接口及其实现块为标准 PLC 逻辑编排
 *                         与诊断镜像层，不构成 ISO 13849 / IEC 62061 认证
 *                         安全功能，安全回路由认证安全控制器/安全 PLC 承载。
 * 契约结构 (Structure)  : 公约 0.11 接口三段式——状态枚举（本文件承载）+
 *                         属性（PROPERTY GET）+ 方法（METHOD）；方法共 4 个
 *                         （≤6 红线内）。故障态一律拒绝方法；门开态下拒绝
 *                         CmdRelock 之外的全部动作。
 * 开源溯源 (Origin)     : 来源标签 tcopen-component / safety-interlock
 *                         （RAW_NOTES_R7 S-2/S-4：TcOpen 组件接口分层思想
 *                         与 ISO 14119 电磁锁扣门联锁公开语义——解锁时序
 *                         状态域、静止确认、审计计数，公开标准资料，仅借
 *                         鉴状态域语义；接口命名、枚举编号、方法签名 100%
 *                         本库独立设计，clean-room 未复制源码）。
 * 归属说明 (Ownership)  : 本文件同时承载 E_DL_SafetyDoorState 枚举定义，该
 *                         枚举归属接口 I_DL_SafetyDoor，与其同文件发布
 *                         （公约 0.11；禁止异文件同名异型重复定义）。
 * 红线自检 (Redline)    : R1 零全局变量表/外部变量引用 ✓｜R2 零物理 IO 地址 ✓
 *                         R3 纯 IEC 61131-3 ✓｜R4 N/A（契约件无运算）
 *                         R5 全成员中英双语同行注释 ✓｜R6 N/A（接口无状态机）
 *                         R7 N/A（无实例调用）｜R18 INTERFACE/END_INTERFACE
 *                         成对终结 ✓
 * 修订历史 (Revision)   :
 *   2026-11-15  v1.0.0  首版入库（Round 07 · DL_Device 安全门族接口件）
 *============================================================================*)

(*-----------------------------------------------------------------------------
 * 枚举: E_DL_SafetyDoorState（归属接口 I_DL_SafetyDoor，与其同文件）
 * 含义: 电磁锁扣门解锁时序离散状态。编号步长 10 留空位，eFault 取 99 保证
 *       排序末位（全库枚举编号惯例）。
 *----------------------------------------------------------------------------*)
TYPE E_DL_SafetyDoorState :
(
    eIdle               := 0,   // 待机：门锁全确认，可受理解锁请求 / Idle, door and lock fully confirmed, unlock acceptable
    eLocked             := 10,  // 已闭锁：关门再锁定确认中或重启抑制保持 / Locked, relock confirming or restart inhibit held
    eStopRequested      := 20,  // 已请求停机：解锁时序中停机请求输出有效 / Stop requested, stop-request output active in the unlock sequence
    eStandstillConfirmed:= 30,  // 静止已确认：零速反馈或 run-down 计时达成 / Standstill confirmed by zero-speed feedback or run-down timer
    eUnlocked           := 40,  // 已解锁：解锁电磁铁输出有效，等待开门 / Unlocked, solenoid energized, awaiting door opening
    eOpened             := 50,  // 门已开启：审计计数已累加，等待关门再锁定 / Opened, audit count incremented, awaiting relock
    eFault              := 99   // 故障锁存：静止超时/防篡改冲突/再锁定超时/非法状态 / Latched fault
) UINT;
END_TYPE

(*-----------------------------------------------------------------------------
 * 接口: I_DL_SafetyDoor
 * 边界防错: 故障态一律拒绝方法并返回 FALSE；门开态下拒绝 CmdRelock 之外的
 *           全部动作；接口层不写物理输出（电磁铁/停机请求由实现块承载）。
 *----------------------------------------------------------------------------*)
INTERFACE I_DL_SafetyDoor

// ---- 属性段（全部只读 GET，实现块一一落地）----------------------------------

PROPERTY eState          : E_DL_SafetyDoorState // 当前解锁时序状态（Current sequence state），枚举见 E_DL_SafetyDoorState
PROPERTY bClosed         : BOOL                 // 门已关闭（Door closed），门关闭反馈镜像 / Door-closed feedback mirror
PROPERTY bLocked         : BOOL                 // 锁已闭锁（Lock engaged），锁闭反馈镜像 / Lock-engaged feedback mirror
PROPERTY bUnlockPermitted: BOOL                 // 允许解锁（Unlock permitted），无故障、无重启抑制且门锁全确认 / Unlock permitted: no fault, no inhibit, door and lock confirmed
PROPERTY bOpened         : BOOL                 // 门开启（Door open），门开启诊断镜像 / Door-open diagnostic mirror
PROPERTY bFault          : BOOL                 // 故障锁存中（Fault latched），显式排除信息级码（R21）/ TRUE = latched fault, info codes excluded
PROPERTY uErrorId        : UDINT                // 末次故障码（Last error code），0=无故障，段位 16#0003_xxxx / Last error code, family 16#0003_xxxx

// ---- 方法段（单发指令，返回受理/合法性结果）----------------------------------

METHOD CmdRequestUnlock : BOOL // 请求解锁（Request unlock）：发起停机请求并进入解锁时序；故障态/门开态拒绝 / Starts the unlock sequence, rejected in fault or door-open
VAR_INPUT
END_VAR

    END_METHOD

METHOD CmdRelock : BOOL // 重新闭锁指令（Relock command）：门开态下关门确认后受理 / Relock, accepted when the door is closed again
VAR_INPUT
END_VAR

    END_METHOD

METHOD CmdReset : BOOL // 复位故障（Reset fault），仅故障态受理返回 TRUE / Reset accepted only in fault state
VAR_INPUT
END_VAR

    END_METHOD

METHOD CmdAuditClear : BOOL // 清除开门审计记录（Clear the open audit count），供批次收尾调用；故障态拒绝 / Clears the open audit count, rejected in fault
VAR_INPUT
END_VAR

    END_METHOD
END_INTERFACE

(* ---- I_DL_StepperOpenLoop.st ---- *)
(*==============================================================================
 * 组件名称 (Component)  : I_DL_StepperOpenLoop
 * 所属子库 (Sublibrary) : DL_Device
 * 当前版本 (Version)    : 1.0.0
 * 分类     (Category)   : 接口（INTERFACE）· 开环步进执行器抽象契约 · Level 1 设备层
 * 作者     (Author)     : Daoli Library
 * 日期     (Date)       : 2026-11-15
 * 兼容性   (Platform)   : CODESYS 3.5 / TwinCAT 3 / 汇川 InoProShop / Schneider
 *                         Machine Expert；纯 IEC 61131-3（第 3 版）接口语法，
 *                         仅依赖 Standard.library，零厂商方言
 * 功能简介 (Function)   : 开环步进电机（脉冲 + 方向型）标准抽象契约。按本库接口
 *                         三段式公约（0.11）组织：配套结构体（组态参数域）+
 *                         属性（PROPERTY GET，只读状态出口）+ 方法（METHOD，
 *                         单发指令入口）。上层工站、手动调试页、HMI 适配层仅
 *                         依赖本接口引用，即可用同一套代码适配脉冲方向型步进
 *                         驱动器、总线型闭环步进（位置模式降级使用）与仿真
 *                         步进轴，实现「契约-实现」分层与零硬件耦合。
 * 方法数红线 (Budget)   : 方法共 6 个，恰在本库接口方法数红线（≤ 6）临界：
 *                         Init / Enable / MoveRelative / Stop / Reset /
 *                         GetErrorId。回原、点动、绝对定位职责不入本接口，
 *                         由上层工艺块以 MoveRelative 组合实现。
 * 开源溯源 (Origin)     : 来源标签 stepper（GitHub topics 开组）+ TcOpen 分层思想。
 *                         仅参考 MIT 许可开源步进驱动项目（AccelStepper 及同类
 *                         公开仓库）的「梯形加减速脉冲频率规划算法思想」与
 *                         「脉冲当量 / 最大速度 / 加速度 / 超时」参数域惯例，
 *                         以及 TcOpen（Apache-2.0）公开的「契约-实现分离 +
 *                         属性/方法三段式」分层范式；本接口的命名、方法签名、
 *                         状态语义与结构体布局 100% 本库独立设计，clean-room
 *                         实现，未复制任何来源的代码行，不构成衍生作品。
 * 归属说明 (Ownership)  : 本文件同时承载 ST_DL_StepperCfg（步进组态结构体），
 *                         该结构体归属接口 I_DL_StepperOpenLoop，与其同文件
 *                         发布（公约 0.18：一文件一 POU + 随宿主发布配套 DUT）。
 *                         状态枚举 E_DL_StepperState 归属实现块
 *                         FB_DL_PulseDirStepper，随其文件发布，本接口不引用。
 * 红线自检 (Redline)    : 全局隔离 ✓（零全局变量表引用、零外部变量声明、零物理
 *                         地址字面记号）｜命名合规 ✓｜注释完整 ✓（结构体成员与
 *                         方法参数 100% 中英双语同行注释）｜OOP 封装 ✓（属性全部
 *                         只读 GET，动作全部经方法受理）｜周期安全 ✓（接口无实例、
 *                         无状态机，方法不驻留跨周期状态）｜防御编程 ✓（契约层
 *                         写死参数域与拒绝语义）｜可移植性 ✓（纯 IEC 61131-3）｜
 *                         终结符成对 ✓（TYPE/END_TYPE、INTERFACE/END_INTERFACE）
 * 设计要点 (Key notes)  : ① 开环本质：fPosition 是「指令推算位置」而非编码器
 *                          反馈位置，接口注释强制声明禁止当反馈用；上层需要真实
 *                          位置必须外挂编码器并另行封装，不得在本接口上做闭环。
 *                         ② 限位与报警经 uAlarmWord 位域统一回读（bit0 正限位 /
 *                          bit1 负限位 / bit2 驱动器报警 / bit3 堵转超时 /
 *                          bit4~15 保留），避免为每类故障各开一个属性。
 *                         ③ 方法返回 FALSE 时 GetErrorId 必须给出非零码，禁止
 *                          静默失败（契约层强制，实现块逐条落地）。
 *                         ④ 方法全部为非阻塞单发语义：方法内只登记请求并置内部
 *                          标志，跨周期动作由实现块主体状态机执行（公约 3.4）。
 * 修订历史 (Revision)   :
 *   2026-11-15  v1.0.0  首版入库（Round 09 · DL_Device 开环步进族 · 契约件）
 *============================================================================*)

(*-----------------------------------------------------------------------------
 * 结构体: ST_DL_StepperCfg（归属接口 I_DL_StepperOpenLoop，与其同文件发布）
 * 用途: 开环步进的机械换算与运动限制参数域。由调用方持有并经 Init 的
 *       VAR_IN_OUT 注入，实现块仅保存副本、不改写调用方数据。
 * 说明: fTaskCycle 字段为 R9 规格字段表之外的增补项（规格实现条款④要求
 *       「脉冲翻转步长由任务周期与频率求导」，而规格字段表未列该字段），
 *       在此留档说明：增补不改变已列字段语义，仅补齐实现所需的周期基准。
 *----------------------------------------------------------------------------*)
TYPE ST_DL_StepperCfg :
STRUCT
    uStepsPerMm  : UINT := 400;        // 脉冲当量（Pulse equivalent）[脉冲/mm]，域 > 0 / Must be greater than zero
    uMicrostep   : UINT := 1;          // 驱动器细分数（Microstep divisor）[细分]，域 >= 1 / Microstep divisor, one or above
    fMaxSpeed    : LREAL := 50.0;      // 最大运行速度（Max travel speed）[mm/s]，域 > 0 / Must be greater than zero
    fAccel       : LREAL := 500.0;     // 加/减速度（Acceleration and deceleration）[mm/s²]，域 > 0 / Symmetric accel and decel, greater than zero
    tStallTimeout : TIME := T#500MS;   // 堵转判据附加裕度（Stall timeout margin）[ms]，叠加在理论耗时之上 / Added on top of the theoretical move time
    fTaskCycle   : LREAL := 0.01;      // 任务周期（Task cycle time）[s]，频率求导与脉冲翻步基准 / Base for frequency derivation and pulse toggling
END_STRUCT
END_TYPE

(*-----------------------------------------------------------------------------
 * 接口: I_DL_StepperOpenLoop
 * 契约结构: 属性（PROPERTY GET）+ 方法（METHOD）两段式；属性 3 个、方法 6 个。
 * 状态跃迁契约（实现块必须逐条保证）：
 *   1 未 Init 或 Init 失败时，除 Enable(FALSE) 与 GetErrorId 外全部方法
 *     返回 FALSE 并置非零码；拒绝路径不得改变任何内部运动状态。
 *   2 Enable(TRUE) 仅在该轴无故障锁存时受理；Enable(FALSE) 恒受理，且必须
 *     在本拍内冻结脉冲输出（不得留半脉冲），偏移/位置保持不清零。
 *   3 MoveRelative 仅在「已使能 + 无故障 + 空闲」时受理；运行中再次调用
 *     必须拒绝（本接口不定义在线改距语义，改距请先 Stop 再下发）。
 *   4 限位触发后 MoveRelative 必须拒绝同方向指令（反方向恒受理，用于脱离
 *     限位）；方向判据为电平判据，不因复位而失效。
 *   5 Stop 为受控停车：按减速度斜坡降频至零后回空闲；故障锁存期间调用
 *     无效（返回 FALSE 并给出码），硬切请用 Enable(FALSE)。
 *   6 Reset 仅在故障锁存时受理；驱动器报警源（uAlarmWord.bit2）未消失时
 *     复位不得真正解除锁存（ADR 口径：报警源优先）。
 *   7 任何跃迁语义变化视为 MAJOR 变更，必须回写子库 VERSION.md 迁移指引。
 *----------------------------------------------------------------------------*)
INTERFACE I_DL_StepperOpenLoop

(* —— 段 1｜属性（PROPERTY GET）：只读状态出口，实现块一一落地 —— *)
PROPERTY bReady      : BOOL  // 就绪（Ready），TRUE = 已初始化 + 已使能 + 无故障 + 空闲 / Initialized, enabled, fault free and idle
PROPERTY fPosition   : LREAL // 指令位置累计（Command position）[mm]，开环推算值，非编码器反馈 / Open-loop derived position, never an encoder feedback
PROPERTY uAlarmWord  : WORD  // 报警字（Alarm word）[bit]：bit0 正限位 / bit1 负限位 / bit2 驱动器报警 / bit3 堵转超时 / bit4~15 保留 / Bit0 positive limit, bit1 negative limit, bit2 drive alarm, bit3 stall timeout, bits 4 to 15 reserved

(* —— 段 2｜方法（METHOD）：单发指令，返回受理结果 —— *)

METHOD Init : BOOL                  // 初始化（Initialize）：注入组态，校验参数域，返回是否成功
VAR_IN_OUT
    stCfg : ST_DL_StepperCfg;       // 步进组态（Stepper configuration），调用方持有，实现块仅存副本 / Caller-owned configuration, the implementation keeps a copy
END_VAR

    END_METHOD

METHOD Enable : BOOL                // 使能/去使能（Enable and disable），电平语义，FALSE 时本拍冻结脉冲
VAR_INPUT
    bEnable : BOOL;                 // 使能指令（Enable command），TRUE = 使能 / FALSE = 去使能并冻结脉冲输出 / TRUE enables, FALSE disables and freezes the pulse output
END_VAR

    END_METHOD

METHOD MoveRelative : BOOL          // 相对位移（Move relative）：从当前指令位置移动指定距离，梯形加减速由实现块规划
VAR_INPUT
    fDistance : LREAL;              // 相对位移（Relative distance）[mm]，正负双向，负值即负向 / Signed distance in millimetres, negative means reverse
    fSpeed    : LREAL;              // 运行速度（Run speed）[mm/s]，域 > 0，超最大速度自动钳位 / Must be positive, clamped to the maximum speed
END_VAR

    END_METHOD

METHOD Stop : BOOL                  // 受控停车（Controlled stop）：按减速度斜坡降频至零并清除当前运动指令
VAR_INPUT
END_VAR

    END_METHOD

METHOD Reset : BOOL                 // 故障复位（Fault reset）：清除限位/堵转/参数类锁存，报警源未消失时不解除
VAR_INPUT
END_VAR

    END_METHOD

METHOD GetErrorId : UDINT           // 故障码查询（Error code query），0 = 无故障；方法返回 FALSE 时必为非零码
VAR_INPUT
END_VAR

    END_METHOD
END_INTERFACE

(* ---- I_DL_TemperatureZone.st ---- *)
(*==============================================================================
 * 组件名称 (Component)  : I_DL_TemperatureZone
 * 所属子库 (Sublibrary) : DL_Device
 * 当前版本 (Version)    : 1.0.0
 * 兼容性   (Platform)   : CODESYS 3.5 / TwinCAT 3 / 汇川 InoProShop / Machine Expert
 *                         纯 IEC 61131-3（第 3 版）OOP 接口契约，零厂商方言
 * 分类     (Category)   : 接口（INTERFACE）· 温控区执行抽象 · Level 1 DL_Device 开库件
 * 功能描述 (Function)   : 加热/冷却温控区标准抽象契约。上层工艺层（炉区、恒温室、
 *                         模温机、老化房）只依赖本接口编程，与具体温控实现
 *                         （FB_DL_HeatCoolZone 等）彻底解耦（依赖倒置）。
 *                         契约按接口三段式公约（0.11）组织：状态枚举 + 只读属性
 *                         （实测温度 / 输出功率 / 状态 / 故障 / 故障码）+ 方法
 *                         （设定值 / 投退 / 复位）；方法共 3 个（红线 ≤6）。
 *                         实现块必须以 IMPLEMENTS 挂接本接口并逐成员兑现。
 * 开源溯源 (Origin)     : 原创设计。状态集合惯例与断偶安全方向语义参考 NAMUR
 *                         NE43 公开标准与温控器行业公知行为（来源标签
 *                         lbp-device / namur-ne43），未参考、未复制任何厂商源码。
 * 本文件内含       : TYPE      E_DL_TempZoneState（状态枚举，归属 DL_Device，
 *                              随本接口同文件发布）
 *                    INTERFACE I_DL_TemperatureZone
 * 依赖     (Depends)    : 无（纯契约文件，零外部引用，可单独编译）
 * 红线自检 (Redline)    : R1 ✓ 零全局变量表与外部变量引用 ｜ R2 ✓ 零物理 IO 地址直写
 *                         R3 ✓ 纯 IEC 61131-3 ｜ R4 ✓ 契约级不适用（无算法分支）
 *                         R5 ✓ 全成员中英双语同行注释 ｜ R6 ✓ 契约级不适用（由实现块承担）
 *                         R7 不适用（无定时器/边沿实例，纯契约）
 * 修订历史 (Revision)   :
 *   2026-11-15  v1.0.0  首版入库 · Round 05 · 泳道 B · 契约出处 ROUND_PLAN_R5 §1.7
 *============================================================================*)

(*-----------------------------------------------------------------------------
 * 枚举: E_DL_TempZoneState（归属 DL_Device，随 I_DL_TemperatureZone 同文件）
 * 含义: 温控区离散状态机。数值步长留空位便于后续插态而不破坏已有工程。
 *----------------------------------------------------------------------------*)
{attribute 'qualified_only'}
{attribute 'strict'}
TYPE E_DL_TempZoneState :
(
    eIdle        := 0,   // 空闲：未投运，双通道切断 / Idle: not commissioned, both channels cut off
    eHeating     := 10,  // 加热中：加热通道输出功率大于热平衡容差 / Heating: heater duty above thermal-balance tolerance
    eCooling     := 20,  // 冷却中：冷却通道输出功率大于热平衡容差 / Cooling: cooler duty above thermal-balance tolerance
    eHolding     := 30,  // 保温中：双通道均处于热平衡容差带内 / Holding: both channels inside thermal-balance tolerance band
    eSensorBreak := 40,  // 断偶锁存：传感器断线/开路，双通道切断待复位 / Sensor break latched: sensor break, channels cut pending reset
    eFault       := 99   // 故障兜底：非法状态或接口引用无效，切断待复位 / Fault fallback: illegal state or invalid interface reference, cut pending reset
) UINT;
END_TYPE

(*-----------------------------------------------------------------------------
 * 接口: I_DL_TemperatureZone
 * 契约说明:
 *   - 属性全部为只读 GET 语义，实现块不得提供 SET 通道（状态只读外泄）。
 *   - 方法均为非阻塞单发语义：方法内只置请求标志，动作由实现块主体状态机
 *     在扫描周期内执行（跨周期动作禁止驻留在方法内部）。
 *   - SetSetpoint 返回值 = 设定值合法性（非有限值一律拒绝并返回 FALSE）。
 *   - CmdReset 返回值 = 当前是否可复位（断偶态要求信号质量恢复后方可成功）。
 *----------------------------------------------------------------------------*)
INTERFACE I_DL_TemperatureZone

// ---- 只读属性段（PROPERTY GET）----------------------------------------------
PROPERTY fTempActual : REAL                 // 实测温度（Actual temperature）[°C]，取自注入的传感器接口
PROPERTY fPowerOut   : REAL                 // 输出功率（Power output）[-100..100 %]，正=加热 / 负=冷却
PROPERTY eState      : E_DL_TempZoneState   // 当前状态机状态（Current zone state）
PROPERTY bFault      : BOOL                 // 故障锁存中（Fault latched），仅故障级状态置位，信息级不置位
PROPERTY uErrorId    : UDINT                // 末次故障/信息码（Last error/info code），0 = 无

// ---- 方法段（METHOD，共 3 个，红线 ≤6）--------------------------------------
METHOD SetSetpoint : BOOL
VAR_INPUT
    fTemp : REAL;                           // 目标温度（Target temperature）[°C]，越界由实现块钳位，非有限值拒绝
END_VAR

    END_METHOD

METHOD CmdEnable
VAR_INPUT
    bOn : BOOL;                             // TRUE=投运（Commission on），FALSE=退出并切断双通道
END_VAR

    END_METHOD

METHOD CmdReset : BOOL                      // 复位故障（Reset fault），返回当前是否可复位
VAR_INPUT
END_VAR

    END_METHOD
END_INTERFACE

(* ---- I_DL_TowerLight.st ---- *)
(*==============================================================================
 * 组件名称 (Component)  : I_DL_TowerLight
 * 所属子库 (Sublibrary) : DL_Device
 * 当前版本 (Version)    : 1.0.0
 * 兼容性   (Platform)   : CODESYS 3.5 / TwinCAT 3 / 汇川 InoProShop / Machine Expert
 *                         纯 IEC 61131-3（第3版）接口语法，零厂商方言
 * 分类     (Category)   : 状态指示抽象接口（Interface）+ 配套枚举 3 个（DUT）
 * 功能描述 (Function)   : 工业安灯塔（Andon 三色/四色塔灯 + 蜂鸣）标准抽象契约。
 *                         按本库接口三段式组织：状态枚举（随文件发布）+ 只读
 *                         属性组（10 个）+ 指令方法组（3 个）。上层 HMI 面板、
 *                         工站顺序控制、PackML 状态机只需持有本接口引用，即可
 *                         适配直驱型（每色一路数字输出）、模块化型（XVU 类
 *                         集束塔灯）与总线型（IO-Link 塔灯）三类实现，而无需
 *                         感知底层通道数量与驱动方式。
 * 接口三段式 (Contract): ①状态枚举：E_DL_TowerColor / E_DL_TowerPattern /
 *                         E_DL_TowerState（均随本文件发布）；②属性：全部只读
 *                         GET（eState / eRed / eAmber / eGreen / eBlue / eWhite /
 *                         bBuzzer / bSilenced / bError / uErrorId 共 10 个）；
 *                         ③方法：SetColor / SilenceBuzzer / Reset 共 3 个，
 *                         满足接口方法不超过 6 个的拆分红线。
 * 边界防错 (Boundary)   : 接口层不做任何电平输出（灯与蜂鸣的物理通道由实现块
 *                         以输出引脚给出）；接口层不读任何现场输入（状态位由
 *                         实现块引脚注入）；红绿互斥属实现块出口断言职责，
 *                         接口只声明属性语义，不承诺仲裁顺序。
 * 开源溯源 (Origin)     : 原创实现（参考 TcOpen 组件范式）。来源标签
 *                         tcopen-component / stack-light（RAW_NOTES_R8 条目 S-13：
 *                         TcOpen 的 stack-light 组件公开文档所呈现的
 *                         「状态位集合 → 灯色仲裁 → 通道输出」三层分层惯例），
 *                         仅借鉴功能分类、接口参数域与状态语义；接口命名、
 *                         属性与方法签名、枚举取值步长按本库红线独立设计，
 *                         clean-room 未复制任何源码行。许可证说明：TcOpen 采用
 *                         MIT 许可，其公开语义描述可自由借鉴；本文件不含其
 *                         任何代码片段，无许可证传染风险。
 * 归属说明 (Ownership)  : 本文件同时承载三个枚举定义，均归属接口
 *                         I_DL_TowerLight，与其同文件发布（公约 0.18：一文件
 *                         一 POU，枚举随宿主发布，禁止在其他文件重复声明）。
 * 验收向量 (Acceptance) : 本文件为纯契约，无执行体，行为验收沿用实现块
 *                         FB_DL_SignalTower 的 V1 至 V8（见该文件头注释）。
 *                         契约级自查三条：C1 属性共 10 个且全部只读 GET；
 *                         C2 方法共 3 个且均带布尔受理返回值；C3 三个枚举取值
 *                         互不重叠且步长为 10，便于后续插值。
 * 已知限制 (Limits)     : 1 eRotate 依赖实现层是否具备环灯硬件，单色通道实现
 *                         退化为慢闪，属实现选择而非契约缺陷。2 接口不约束仲裁
 *                         优先序与通道数量，跨实现的行为一致性由各实现块头注释
 *                         的优先级表承担。3 消音权限与消音次数限制属上层 HMI
 *                         职责，不在本契约内。
 * 规格偏离 (R11 Dev.)   : 无。三个枚举取值、10 个属性类型与 3 个方法签名与
 *                         规格第 3.1 节逐条一致。
 * 红线自检 (Redline)    : 零全局变量表访问 ✓｜零外部变量声明 ✓｜零物理地址直写 ✓
 *                         纯 IEC 61131-3 ✓｜全成员中英双语同行注释 ✓
 *                         INTERFACE 与 END_INTERFACE 成对 ✓｜三个 TYPE 与 END_TYPE 成对 ✓
 * 修订历史 (Revision)   :
 *   2026-11-15  v1.0.0  首版入库（Round 08 · 泳道 C · DL_Device 状态指示族）
 *============================================================================*)

(*-----------------------------------------------------------------------------
 * 枚举: E_DL_TowerColor（归属接口 I_DL_TowerLight，与其同文件）
 * 含义: 塔灯灯色通道。数值步长 10 留空位，便于后续插入特殊色（如紫色、
 *       青色）而不破坏已有工程持久化的数值。
 *----------------------------------------------------------------------------*)
TYPE E_DL_TowerColor :
(
    eNone  := 0,     // 无色 / 清除该色通道（No color, channel cleared）
    eRed   := 10,    // 红色（Red），安全与未确认故障主色，优先级最高
    eAmber := 20,    // 黄色 / 琥珀色（Amber），预警与待处理主色
    eGreen := 30,    // 绿色（Green），自动运行正常主色
    eBlue  := 40,    // 蓝色（Blue），手动模式与操作员求助主色
    eWhite := 50     // 白色（White），待机与就绪指示（可选通道）
) UINT;
END_TYPE

(*-----------------------------------------------------------------------------
 * 枚举: E_DL_TowerPattern（归属接口 I_DL_TowerLight，与其同文件）
 * 含义: 单色通道的显示模式。闪烁时基一律由实现块的半周期引脚给定，
 *       禁止读取任何内部时钟源。
 *----------------------------------------------------------------------------*)
TYPE E_DL_TowerPattern :
(
    eOff        := 0,   // 熄灭（Off），该色通道无输出
    eSteady     := 10,  // 常亮（Steady），电平恒为真
    eFlashSlow  := 20,  // 慢闪（Slow flash），默认半周期 500 毫秒，全周期约 1 赫兹
    eFlashFast  := 30,  // 快闪（Fast flash），默认半周期 250 毫秒，全周期约 2 赫兹
    eRotate     := 40   // 旋转（Rotate），多色环灯逐色轮转；单色通道实现退化为慢闪
) UINT;
END_TYPE

(*-----------------------------------------------------------------------------
 * 枚举: E_DL_TowerState（归属接口 I_DL_TowerLight，与其同文件）
 * 含义: 塔灯"显示状态"的语义分类，取值为仲裁结果的唯一出口分类，不是
 *       实现块内部私有步序；上层可据此做 HMI 文本映射与报警分级。
 *----------------------------------------------------------------------------*)
TYPE E_DL_TowerState :
(
    eNormal      := 0,   // 正常 / 待机（Normal or standby），无主级告警
    eWarning     := 10,  // 预警（Warning），未确认慢闪、已确认常亮
    eFaultAck    := 20,  // 故障已确认（Fault acknowledged），红常亮不鸣
    eFaultUnack  := 30,  // 故障未确认（Fault unacknowledged），红慢闪并鸣
    eSafety      := 40,  // 安全事件（Safety event），红快闪强制鸣，最高优先
    eManual      := 50,  // 手动模式（Manual mode），蓝常亮
    eCall        := 60   // 操作员求助（Operator call），蓝快闪
) UINT;
END_TYPE

(*-----------------------------------------------------------------------------
 * 接口: I_DL_TowerLight
 * 契约结构: 属性（只读 GET，10 个）+ 方法（3 个）两段式，方法总数满足
 *           不超过 6 个的拆分红线。方法均为非阻塞单发语义，不含跨扫描周期
 *           状态驻留；返回值仅表示"请求是否被受理"，实际灯效以属性为准。
 * 受理语义: SetColor 在更高优先级占用或故障锁存时返回 FALSE；
 *           SilenceBuzzer 在非蜂鸣期或安全事件期返回 FALSE（安全事件不受
 *           消音约束）；Reset 仅在存在故障锁存时返回 TRUE。
 *----------------------------------------------------------------------------*)
INTERFACE I_DL_TowerLight

// ---- 属性段（全部只读 GET，共 10 个）--------------------------------------

PROPERTY eState     : E_DL_TowerState   // 当前显示状态（Displayed state），等于仲裁结果的语义分类
PROPERTY eRed       : E_DL_TowerPattern // 红色通道当前模式（Red pattern），eOff=不亮
PROPERTY eAmber     : E_DL_TowerPattern // 黄色通道当前模式（Amber pattern），eOff=不亮
PROPERTY eGreen     : E_DL_TowerPattern // 绿色通道当前模式（Green pattern），eOff=不亮
PROPERTY eBlue      : E_DL_TowerPattern // 蓝色通道当前模式（Blue pattern），eOff=不亮
PROPERTY eWhite     : E_DL_TowerPattern // 白色通道当前模式（White pattern），eOff=不亮
PROPERTY bBuzzer    : BOOL              // 蜂鸣器当前输出（Buzzer active），TRUE=正在鸣响
PROPERTY bSilenced  : BOOL              // 已消音（Silenced），消音保持窗内为 TRUE
PROPERTY bError     : BOOL              // 故障锁存（Fault latched），仅故障级码置位，信息级码不置位
PROPERTY uErrorId   : UDINT             // 错误码（Error code），0=无错误，段位 16#0003_xxxx

// ---- 方法段（单发指令，返回受理结果，共 3 个）-----------------------------

(* 请求置某色某模式（Set color and pattern）；返回 FALSE 表示当前被更高优先级
 * 占用、处于故障锁存或使能关闭。色通道生命周期由实现块仲裁表裁决。 *)
METHOD SetColor : BOOL
VAR_INPUT
    eColor   : E_DL_TowerColor;    // 目标灯色（Target color），eNone=撤销人工覆盖
    ePattern : E_DL_TowerPattern;  // 目标模式（Target pattern），eOff=该色熄灭
END_VAR

(* 消音（Silence buzzer）：一次性受理，超过保持时长自动恢复蜂鸣；非蜂鸣期或
 * 处于安全事件期返回 FALSE（安全事件不受消音约束）。 *)
    END_METHOD

METHOD SilenceBuzzer : BOOL
VAR_INPUT
END_VAR

(* 复位故障锁存（Reset fault latch）：仅存在锁存故障时返回 TRUE，否则 FALSE。 *)
    END_METHOD

METHOD Reset : BOOL
VAR_INPUT
END_VAR

    END_METHOD
END_INTERFACE

(* ---- I_DL_VacuumGenerator.st ---- *)
(*==============================================================================
 * 组件名称 (Component)  : I_DL_VacuumGenerator
 * 所属子库 (Sublibrary) : DL_Device
 * 当前版本 (Version)    : 1.0.0
 * 兼容性   (Platform)   : CODESYS 3.5 / TwinCAT 3 / 汇川 InoProShop / Machine Expert
 *                         纯 IEC 61131-3（第3版）接口语法，零厂商方言
 * 分类     (Category)   : 设备抽象接口（Interface）+ 配套状态枚举（DUT）
 * 功能简述 (Function)   : 真空发生器（负压吸盘供气）标准抽象契约。定义状态
 *                         读取属性组（GET）与真空建立/破真空/停止/复位方法
 *                         组，供 DL_Process 拾放工站（PickAndPlaceStation /
 *                         CellFeederVacuum）做依赖注入与解耦调用；具体电磁
 *                         阀驱动、负压采集与吹气脉冲由实现块（如
 *                         FB_DL_VacuumEjector）完成，接口层不做任何过程
 *                         映像读写，仅承载纯软件契约。
 * 开源溯源 (Origin)     : 来源标签 lbp-device（RAW_NOTES_R6 S-1：真空吸拾
 *                         放的建立-保持-破真空三段操作惯例、负压域压力
 *                         反馈语义等行业公知工程惯例，公开教学资料，仅借鉴
 *                         通用工程语义；接口命名、方法签名按本库红线独立
 *                         设计，clean-room 未复制源码）。
 * 红线自检 (Redline)    : R1 零全局变量表/外部变量引用 ✓｜R2 零物理 IO 地址 ✓
 *                         R3 纯 IEC 61131-3 ✓｜R5 全成员中英双语同行注释 ✓
 *                         R18 接口以 END_INTERFACE 成对终结 ✓
 * 归属说明 (Ownership)  : 本文件同时承载 E_DL_VacuumState 枚举定义，该枚举
 *                         归属接口 I_DL_VacuumGenerator，与其同文件发布。
 * 修订历史 (Revision)   :
 *   2026-11-15  v1.0.0  首版入库（R6 轮 · DL_Device 阀门/驱动族深化）
 *============================================================================*)

(*-----------------------------------------------------------------------------
 * 枚举: E_DL_VacuumState（归属接口 I_DL_VacuumGenerator，与其同文件）
 * 含义: 真空发生器状态机离散状态。数值步长 10 留空位，便于后续插态
 *       而不破坏已有工程的持久化数值；eFault 取 99 保证排序末位。
 *----------------------------------------------------------------------------*)
TYPE E_DL_VacuumState :
(
    eIdle       := 0,    // 空闲稳态：双阀全断，不吸附不吹气 / Idle steady state, both valves off, no evacuate or blow-off
    eEvacuating := 10,   // 抽真空中：真空阀开，等待负压建立确认 / Evacuating, vacuum valve open, awaiting vacuum establishment confirmation
    eVacuumOk   := 20,   // 真空建立确认：负压阈值（及可选开关）确认的吸附保持态 / Vacuum established, holding state confirmed by threshold and optional switch
    eBlowing    := 30,   // 破真空吹气中：吹气阀定宽脉冲输出，真空阀强制断 / Blowing, blow-off valve in fixed-width pulse, vacuum valve forced off
    eFault      := 99    // 故障锁存态：超时/反馈失效/非法状态，仅复位可清 / Latched fault state (timeout, feedback loss), cleared only by reset
) UINT;
END_TYPE

(*-----------------------------------------------------------------------------
 * 接口: I_DL_VacuumGenerator
 * 契约结构: 属性（PROPERTY GET）+ 方法（METHOD）两段式；方法总数 4 个，
 *           满足接口方法 ≤6 的拆分红线。所有方法均为非阻塞单发语义，
 *           不含跨扫描周期状态驻留；返回值仅表示"指令是否被受理"，
 *           实际真空状态以属性 eState/bVacuumOk 为准。
 * 边界防错: 任何动作方法在故障锁存态一律拒绝并返回 FALSE；实现块负责
 *           阀输出与负压采集的全部过程映像交互，本接口不涉及。
 *----------------------------------------------------------------------------*)
INTERFACE I_DL_VacuumGenerator

// ---- 属性段（全部只读 GET）------------------------------------------------

PROPERTY eState    : E_DL_VacuumState // 当前状态机状态（Current state）
PROPERTY bVacuumOk : BOOL             // 真空建立确认（Vacuum established），TRUE=吸附保持中 / TRUE = vacuum established and holding
PROPERTY fPressure : REAL             // 负压反馈值（Pressure feedback）[kPa]，0=大气压，负值=真空度 / Pressure feedback [kPa], 0 = atmospheric, negative = vacuum
PROPERTY bFault    : BOOL             // 故障锁存中（Fault latched），TRUE=存在未复位故障 / TRUE = latched fault present
PROPERTY uErrorId  : UDINT            // 末次故障码（Last error code），0=无故障，段位 16#0003_xxxx / Last error code, 0 = none, family 16#0003_xxxx

// ---- 方法段（单发指令，返回受理结果）--------------------------------------

METHOD CmdEvacuate : BOOL // 建立真空指令（Evacuate command），单发；故障态拒绝返回 FALSE / Rejected with FALSE in fault state
VAR_INPUT
END_VAR

    END_METHOD

METHOD CmdBlowOff : BOOL // 破真空吹气指令（Blow-off command），单发，实现块输出定宽脉冲 / One-shot blow-off, fixed-width pulse by implementation
VAR_INPUT
END_VAR

    END_METHOD

METHOD CmdStop : BOOL // 双阀全断保持现状（Stop command, both valves off, hold state）；故障态拒绝返回 FALSE / Rejected with FALSE in fault state
VAR_INPUT
END_VAR

    END_METHOD

METHOD CmdReset : BOOL // 复位指令（Reset command），返回是否可复位（存在故障时为 TRUE）/ Returns TRUE only when resettable
VAR_INPUT
END_VAR

    END_METHOD
END_INTERFACE

(* ---- I_DL_VfdDrive.st ---- *)
(*==============================================================================
 * 组件名称 (Component)  : I_DL_VfdDrive
 * 所属子库 (Sublibrary) : DL_Device
 * 当前版本 (Version)    : 1.0.0
 * 兼容性   (Platform)   : CODESYS 3.5 / TwinCAT 3 / 汇川 InoProShop / Machine Expert
 *                         纯 IEC 61131-3（第3版）接口语法，零厂商方言
 * 分类     (Category)   : 设备抽象接口（Interface）+ 配套状态枚举（DUT）
 * 功能简述 (Function)   : 通用变频器抽象契约（端子型/通信型均可适配）。
 *                         定义状态读取属性组（GET）与运行/停止/点动/频率
 *                         设定/多段速选择/复位方法组，供风机泵类与输送线
 *                         驱动层做依赖注入与解耦调用；端子输出、模拟量
 *                         给定与反馈采集由实现块（如 FB_DL_VfdGeneric）
 *                         完成，接口层不做任何过程映像读写。
 * 开源溯源 (Origin)     : 来源标签 lbp-basic-process / lbp-device
 *                         （RAW_NOTES_R6 S-1 + S-4：变频器控制标准信号集
 *                         ——运行/正反转/点动/多段速/频率到达/故障复位
 *                         端子语义，公开技术资料，仅借鉴通用信号域语义；
 *                         接口命名、方法签名按本库红线独立设计，clean-room
 *                         未复制源码）。
 * 红线自检 (Redline)    : R1 零全局变量表/外部变量引用 ✓｜R2 零物理 IO 地址 ✓
 *                         R3 纯 IEC 61131-3 ✓｜R5 全成员中英双语同行注释 ✓
 *                         R18 接口以 END_INTERFACE 成对终结 ✓
 * 归属说明 (Ownership)  : 本文件同时承载 E_DL_VfdState 枚举定义，该枚举
 *                         归属接口 I_DL_VfdDrive，与其同文件发布。
 * 修订历史 (Revision)   :
 *   2026-11-15  v1.0.0  首版入库（R6 轮 · DL_Device 阀门/驱动族深化）
 *============================================================================*)

(*-----------------------------------------------------------------------------
 * 枚举: E_DL_VfdState（归属接口 I_DL_VfdDrive，与其同文件）
 * 含义: 变频器状态机离散状态。数值步长 10 留空位，便于后续插态
 *       而不破坏已有工程的持久化数值；eFault 取 99 保证排序末位。
 *----------------------------------------------------------------------------*)
TYPE E_DL_VfdState :
(
    eDisabled    := 0,    // 未使能态：驱动未上电/未使能，全部输出切断 / Disabled, drive not enabled, all outputs cut off
    eReady       := 10,   // 就绪态：使能完成，等待运行/点动指令 / Ready, enabled and awaiting run or jog commands
    eRunningFwd  := 20,   // 正转运行态：正转端子输出有效 / Running forward, forward terminal active
    eRunningRev  := 30,   // 反转运行态：反转端子输出有效 / Running reverse, reverse terminal active
    eJogging     := 40,   // 点动态：点动端子输出有效，优先级高于运行 / Jogging, jog terminal active with priority over run
    eFault       := 99    // 故障锁存态：驱动故障/反馈超时/非法状态，复位脉冲可尝试恢复 / Latched fault state (drive fault, feedback timeout), reset pulse may recover
) UINT;
END_TYPE

(*-----------------------------------------------------------------------------
 * 接口: I_DL_VfdDrive
 * 契约结构: 属性（PROPERTY GET）+ 方法（METHOD）两段式；方法总数 6 个，
 *           达接口方法 ≤6 拆分红线的临界值。所有方法均为非阻塞单发
 *           语义，不含跨扫描周期状态驻留；返回值仅表示"指令是否被
 *           受理/参数是否合法"，实际运行状态以属性 eState/bRunning
 *           为准。
 * 边界防错: 故障态下运行/点动/设定类方法一律拒绝并返回 FALSE；复位
 *           方法返回是否受理；实现块负责端子输出与反馈采集的全部
 *           过程映像交互，本接口不涉及。
 *----------------------------------------------------------------------------*)
INTERFACE I_DL_VfdDrive

// ---- 属性段（全部只读 GET）------------------------------------------------

PROPERTY eState       : E_DL_VfdState // 当前状态机状态（Current state）
PROPERTY fFreqSetpoint : REAL         // 频率设定（Frequency setpoint）[Hz]，钳位后生效值 / Effective frequency setpoint [Hz] after clamping
PROPERTY fFreqActual  : REAL          // 频率反馈（Frequency feedback）[Hz]，非有限值时保持末次有效值 / Frequency feedback [Hz], holds last valid on non-finite input
PROPERTY bRunning     : BOOL          // 运行反馈（Running feedback），正转/反转/点动态输出运行中 / TRUE while running forward/reverse or jogging
PROPERTY bFault       : BOOL          // 故障锁存中（Fault latched），TRUE=存在未复位故障 / TRUE = latched fault present
PROPERTY uErrorId     : UDINT         // 末次故障码（Last error code），0=无故障，段位 16#0003_xxxx / Last error code, 0 = none, family 16#0003_xxxx

// ---- 方法段（单发指令，返回受理/合法性结果）--------------------------------

METHOD CmdRun : BOOL // 正/反转运行指令（Run command，bFwd=TRUE 正转 / FALSE 反转），电平语义受理为保持锁存；故障态拒绝返回 FALSE / Run command, held latch accepted, rejected in fault
VAR_INPUT
    bFwd : BOOL; // 方向选择（Direction select），TRUE=正转 / FALSE=反转 / TRUE = forward, FALSE = reverse
END_VAR

    END_METHOD

METHOD CmdStop : BOOL // 停止指令（Stop command）：撤销运行/点动锁存；无条件受理 / Stop command, revokes run and jog latches, unconditionally accepted
VAR_INPUT
END_VAR

    END_METHOD

METHOD CmdJog : BOOL // 点动指令（Jog command，bFwd=TRUE 正向点动），优先级高于运行；故障态拒绝返回 FALSE / Jog command with priority over run, rejected in fault
VAR_INPUT
    bFwd : BOOL; // 点动方向（Jog direction），TRUE=正向 / FALSE=撤销点动保持 / TRUE = jog forward, FALSE = release jog hold
END_VAR

    END_METHOD

METHOD SetFrequency : BOOL // 频率设定（Frequency set）[Hz]，越界/非有限值拒绝并返回 FALSE / Frequency set command, out-of-range or non-finite returns FALSE
VAR_INPUT
    fHz : REAL; // 频率设定值（Frequency value）[Hz]，域 0..fFreqMax / Frequency value [Hz], range 0..fFreqMax
END_VAR

    END_METHOD

METHOD SelectPresetSpeed : BOOL // 多段速选择（Preset speed select），0=模拟量给定、1..7=段速；越界拒绝返回 FALSE / Preset speed select, 0 = analog reference, 1..7 = preset steps, out-of-range returns FALSE
VAR_INPUT
    nIdx : USINT; // 段速索引（Preset index），0=模拟量给定 / 1..7=段速 / Preset index, 0 = analog reference, 1..7 = preset steps
END_VAR

    END_METHOD

METHOD CmdReset : BOOL // 复位指令（Reset command），返回是否受理（存在故障时为 TRUE）/ Returns TRUE only when accepted
VAR_INPUT
END_VAR

    END_METHOD
END_INTERFACE

(* ---- ST_DL_EtSlaveDiagBase.st ---- *)
// ST_DL_EtSlaveDiagBase v1.0.0
// 开源溯源：TcOpen / URL https://github.com/TcOpenGroup / 许可证 MIT / 借鉴 EtcSlaveBase 结构语义（从站诊断基），clean-room 重写
(*
  道莅工业代码库 | DL_Device | ST_DL_EtSlaveDiagBase
  版本: 1.0.0 | 日期: 2026-11-23 | 轮次: R75
  功能: EtherCAT 从站诊断基结构（AL 状态/在线/DC 同步/错误计数字段聚合），
        供各品牌从站诊断 FB 组合扩展
  邻件关系: 与 ProfinetAlarmDiag（PROFINET 告警诊断）协议域不同；本件为
            EtherCAT 域首件结构属主；同步单元级诊断见 ST_DL_EtSyncUnitDiagBase
            （设备级 vs 单元级聚合）
  命名声明: clean-room 重构，字段名全为自命名语义名，不含任何厂商库
            哈希后缀名（原队列条目 EtcSlaveBase_82538BE2 语义对标）
*)
TYPE ST_DL_EtSlaveDiagBase :
STRUCT
    uSlaveAddr      : UINT;      // 从站物理地址 [站号] / EtherCAT slave physical address
    bSlaveOnline    : BOOL;      // 从站在线标志 [-] / Slave online flag
    bSlavePresent   : BOOL;      // 从站配置存在（扫描表匹配）[-] / Slave present per scan list match
    nAlState        : USINT;     // AL 状态码 [码值，0=Init..8=Op] / AL state code, 0=Init..8=Op
    nAlErrCode      : UINT;      // AL 错误码 [AL status code] / AL error status code
    bDcSyncOk       : BOOL;      // 分布式时钟同步合格 [-] / Distributed clock sync ok
    nDcDiffUs       : DINT;      // DC 偏差 [微秒 us] / DC deviation [us]
    uWcStateCnt     : UDINT;     // 工作计数器读数 [计数] / Working counter reading
    uErrFrameCnt    : UDINT;     // 错误帧累计 [帧] / Error frame cumulative count
    uLostLinkCnt    : UDINT;     // 链路丢失累计 [次] / Lost link cumulative count
    bDiagStale      : BOOL;      // 诊断数据过期（看门狗超时）[-] / Diagnostic data stale flag
END_STRUCT
END_TYPE

(* ---- ST_DL_EtSyncUnitDiagBase.st ---- *)
// ST_DL_EtSyncUnitDiagBase v1.0.0
// 开源溯源：TcOpen / URL https://github.com/TcOpenGroup / 许可证 MIT / 借鉴 SyncUnitsBase 结构语义（同步单元诊断基），clean-room 重写
(*
  道莅工业代码库 | DL_Device | ST_DL_EtSyncUnitDiagBase
  版本: 1.0.0 | 日期: 2026-11-23 | 轮次: R75
  功能: EtherCAT 同步单元（Sync Unit）诊断基结构（单元号/参考时钟/成员
        从站索引表/同步质量聚合），供任务级同步诊断 FB 组合扩展
  邻件关系: 与 ST_DL_EtSlaveDiagBase（本批 S10）同族 —— 差异点：从站件为
            单站设备级字段，本件为多站单元级聚合（成员索引表 + 单元级
            同步质量），两件互不嵌套、平级组合
  命名声明: clean-room 重构，不含厂商库哈希后缀名（原队列条目
            SyncUnitsBase_AD6C35CE 语义对标）
*)
TYPE ST_DL_EtSyncUnitDiagBase :
STRUCT
    uSyncUnitId     : UINT;      // 同步单元编号 [单元号] / Sync unit identifier
    bUnitActive     : BOOL;      // 单元激活标志 [-] / Unit active flag
    bRefClockOk     : BOOL;      // 参考时钟锁定 [-] / Reference clock locked
    bAllInSync      : BOOL;      // 全成员同步合格 [-] / All members in sync
    nMemberCnt      : INT;       // 成员从站数 [个]，域 0..8 / Member slave count, domain 0..8
    aMemberAddr     : ARRAY[1..8] OF UINT;   // 成员从站地址表 [站号] / Member slave address table
    nWorstDiffUs    : DINT;      // 成员最大 DC 偏差 [微秒 us] / Worst member DC deviation [us]
    uSyncErrCnt     : UDINT;     // 单元同步错误累计 [次] / Unit sync error cumulative count
    uCycleMissCnt   : UDINT;     // 周期帧丢失累计 [次] / Cycle frame miss cumulative count
    bDiagStale      : BOOL;      // 诊断数据过期（看门狗超时）[-] / Diagnostic data stale flag
END_STRUCT
END_TYPE

(* ---- I_DL_Gripper.st ---- *)
(*
    I_DL_Gripper —— 平行夹爪契约
    ------------------------------------------------------------------
    分类      : DL_Device / Actuator
    前缀      : I_DL_
    版本      : 1.0.0
    溯源      : T2-6 Rockwell AOI（只借「设备级 AOI 粒度 = 阀 / 电机 / 夹爪三件套」
                这一分类事实）；T1-5 开源契约-实现分离范式（Apache-2.0 公开资料，
                仅借分层思想）；方法签名、属性集合、枚举引用 100% 自有；
                clean-room 重写，未复制任何闭源厂商源码，参考实现仅限 MIT/Apache 许可
    平台      : 纯 IEC 61131-3（第3版）接口语法，CODESYS V3.5+ / TwinCAT 3 / InoProShop 通用
    作者      : 道莅代码库 · PLC编程专家（R18）
    ------------------------------------------------------------------
    功能说明  : 把「夹爪」的对外能力收敛为 7 个只读属性加 4 个方法，实现类可换电动 /
                气动 / 伺服夹爪而工艺层零改动（面向接口编程，依赖注入）；
                方法均为一发即走的单发语义，结果经属性回读，方法内部不含跨扫描周期
                状态驻留（跨周期动作在实现块主体完成）；
                ClearFault 只清锁存，绝不隐式产生动作——热复位必须先排除物理原因；
                职责边界：本件只是契约，不采集信号、不驱动电磁阀，全部实现归
                FB_DL_ParallelGripper。
    错误码    : 本件为接口契约，无实现无码位；码位见 FB_DL_ParallelGripper
                （族内 5 槽 16#0003_0166 / 0167 / 032A / 032B / 032C 全部归实现件）
    码位总账  : 不占码位（接口件），实现件码位见 16#0003_0166 / 16#0003_0167 / 16#0003_032A / 16#0003_032B / 16#0003_032C
    状态机    : N/A —— 接口无实现体，状态机归实现件（E_DL_GripperState 随实现件发布）
    采样约定  : 接口不含时间量；实时性由实现件在其所在任务中承担
    修订记录  : 2026-11-16 v1.0.0 首次入库（R18）
*)

(*-----------------------------------------------------------------------------
 * 接口: I_DL_Gripper
 * 契约结构: 只读属性段（GET，7 个）+ 方法段（4 个）
 * 方法数约束: 4 个，满足接口方法不超过 6 个的拆分红线（职责未过载）
 * 边界防错: 故障锁存期间动作方法一律拒绝；ClearFault 只清锁存不产生动作；
 *           eHealth 引用库内唯一属主枚举 E_DL_Ne107Status，本件不重声明（R13 纪律）
 *----------------------------------------------------------------------------*)
INTERFACE I_DL_Gripper

// ---- 属性段（全部只读 GET）------------------------------------------------

PROPERTY bOpened           : BOOL              // 全开到位 / fully opened
PROPERTY bClosed           : BOOL              // 闭合到位（含夹持工件）/ fully closed, the workpiece clamped
PROPERTY bWorkpiecePresent : BOOL              // 工件在位（工件检测信号）/ workpiece present, from the part sensor
PROPERTY fWidth            : REAL              // 当前开口宽度 [mm] / current opening width [mm]
PROPERTY eHealth           : E_DL_Ne107Status  // 健康状态，引用库内唯一属主枚举 / health state, referencing the single owner enum
PROPERTY uErrorId          : UDINT             // 末次故障码，0 = 无故障，段位 16#0003_ / last error code, 0 = none, family 16#0003_
PROPERTY bError            : BOOL              // 故障锁存中，TRUE = 存在未复位故障 / fault latched, TRUE means an unrecovered fault exists

// ---- 方法段（单发指令，结果经属性回读）------------------------------------

METHOD Open : BOOL                             // 请求张开，到位由 bOpened 反映 / request opening, arrival is reflected by bOpened
VAR_INPUT
END_VAR

    END_METHOD

METHOD Close : BOOL                            // 请求闭合到指定夹持力 / request closing at the given clamping force
VAR_INPUT
    fForceSetpoint : REAL;                     // 目标夹持力 [%]，范围 0.0~100.0 / target clamping force [%], range 0.0~100.0
END_VAR

    END_METHOD

METHOD Release : BOOL                          // 松开并撤力，区别于 Open：不放到位只泄力 / release and drop the force, unlike Open it does not drive to the open end
VAR_INPUT
END_VAR

    END_METHOD

METHOD ClearFault : BOOL                       // 清故障锁存（热复位），不产生任何动作 / clear the fault latch, produces no motion
VAR_INPUT
END_VAR

    END_METHOD
END_INTERFACE

(* ---- FC_DL_AisleLeakageMixCalc.st ---- *)
(*
 * FC_DL_AisleLeakageMixCalc | C2 | DL_Device
 * 功能：冷热通道旁通泄漏的混合温度与冷量损失温差       单位：温度 [℃]、泄漏比例 [1]、温差 [K]
 * 工况边界：线性混合模型（无相变、无风机温升），适用于同一机房冷热通道压差稳定的场合；泄漏比例按 [0,1] 物理域钳位，越界仅置信息位（判据取自未钳位原值，R5/R24）；温度须有限
 * 代数值回代：cold=22、hot=35、leak=0.15 → Tmix=0.15×35+0.85×22=23.95 ℃；冷量损失温差=23.95−22=1.95 K（与 spec 回代行一致）
 * 开源溯源：clean-room 自研，未复制任何第三方代码（无外部来源）
 *)
FUNCTION FC_DL_AisleLeakageMixCalc : BOOL
VAR_INPUT
    rColdC     : REAL := 22.0;       // 冷通道送风温度 | cold aisle supply temperature [℃]
    rHotC      : REAL := 35.0;       // 热通道回风温度 | hot aisle return temperature [℃]
    rLeakRatio : REAL := 0.15;       // 旁通泄漏比例 | bypass leakage ratio [1]
END_VAR
VAR_OUTPUT
    rMixedC            : REAL;       // 混合后进柜温度 | mixed rack inlet temperature [℃]
    rColdSupplyDeficitK: REAL;       // 冷量损失温差（混合−冷通道）| cooling loss temperature difference [K]
    rLeakUsed          : REAL;       // 实际参与计算的泄漏比例（已钳位）| leakage ratio actually used, clamped [1]
    xLeakClamped       : BOOL;       // 泄漏比例越界被钳位（信息级）| ratio out of range and clamped, informational
    xValid             : BOOL;       // 输出有效 | outputs valid
END_VAR
VAR
    xFinC : BOOL;                    // 冷通道温度有限性 | cold aisle temperature is finite
    xFinH : BOOL;                    // 热通道温度有限性 | hot aisle temperature is finite
    xFinL : BOOL;                    // 泄漏比例有限性 | leakage ratio is finite
END_VAR
VAR CONSTANT
    DL_ALM_RATIO_LO : REAL := 0.0;   // 泄漏比例下限 | leakage ratio lower bound [1]
    DL_ALM_RATIO_HI : REAL := 1.0;   // 泄漏比例上限 | leakage ratio upper bound [1]
END_VAR

// 段1｜非有限闸（R19）
xFinC := (rColdC = rColdC) AND ((rColdC - rColdC) = 0.0);
xFinH := (rHotC = rHotC) AND ((rHotC - rHotC) = 0.0);
xFinL := (rLeakRatio = rLeakRatio) AND ((rLeakRatio - rLeakRatio) = 0.0);
IF (NOT xFinC) OR (NOT xFinH) OR (NOT xFinL) THEN
    rMixedC := 0.0;                  // 安全值：混合温度 0（下游按无效丢弃）| safe value, downstream discards it
    rColdSupplyDeficitK := 0.0;
    rLeakUsed := 0.0;
    xLeakClamped := FALSE;
    xValid := FALSE;
    FC_DL_AisleLeakageMixCalc := FALSE;
    RETURN;
END_IF

// 段2｜域钳位：泄漏比例物理域 [0,1]，越界标志取自未钳位原值（R24）
IF rLeakRatio < DL_ALM_RATIO_LO THEN
    xLeakClamped := TRUE;
    rLeakUsed := DL_ALM_RATIO_LO;
ELSIF rLeakRatio > DL_ALM_RATIO_HI THEN
    xLeakClamped := TRUE;
    rLeakUsed := DL_ALM_RATIO_HI;
ELSE
    xLeakClamped := FALSE;
    rLeakUsed := rLeakRatio;
END_IF

// 段3｜算法：Tmix = leak×hot + (1−leak)×cold
rMixedC := rLeakUsed * rHotC + (1.0 - rLeakUsed) * rColdC;
rColdSupplyDeficitK := rMixedC - rColdC;

// 段4｜出口
xValid := TRUE;
FC_DL_AisleLeakageMixCalc := TRUE;
END_FUNCTION

(* ---- FC_DL_AnalyzerRecalDaysCalc.st ---- *)
(* ============================================================
   DL_Device / FC_DL_AnalyzerRecalDaysCalc ｜ v1.0.0 ｜ 2026-11-25
   功能：距重新标定天数 nDays = (fDriftLimit − |fDriftNow|) / |fDriftRate| − 已标定天数，
         已标定天数由 tSinceCal 折算（1 天 = 86400 s = 8.64E7 ms）。负值即已超标。
   边界：|fDriftRate| ≤ 1E-9 → 返回哨兵 32767 天、bOverdue=FALSE（永不超期，防除零）；
         允许漂移上限 ≤ 0 → 天数 0、bOverdue=TRUE（组态非法按已超期，安全侧）；
         任一浮点入参非有限 → 天数 0、bOverdue=TRUE（N1）；
         实数转 INT 前先钳到 ±32000（R151：防溢出导致方向翻转）。
         量纲清单（N5）：fDriftRate 为「标定单位/天」，与 fDriftLimit、fDriftNow 同量纲；
         1 天 = 86400 s；TIME_TO_REAL 返回 [ms]，故天数 = ms / 1000 / 86400。
   依赖：仅 IEC 61131-3（ABS / TIME_TO_REAL / REAL_TO_INT） ｜ 溯源：DLF-D-WATERANA
   验收：limit=2.0、now=0.5、rate=0.05/天、已过 10 天 → 1.5/0.05 − 10 = 20 天、FALSE；
         rate=0 → 32767 天；now=2.5 → 负值且 bOverdue=TRUE。
   ============================================================ *)
FUNCTION FC_DL_AnalyzerRecalDaysCalc : BOOL
VAR_INPUT
    fDriftRate  : REAL;  // 漂移速率（标定单位/天，符号无关）[单位/天] / Drift rate per day
    fDriftLimit : REAL;  // 允许总漂移上限 [单位] / Allowed total drift
    fDriftNow   : REAL;  // 当前累计漂移 [单位] / Current accumulated drift
    tSinceCal   : TIME;  // 距上次标定的时长 [ms] / Elapsed time since the last calibration
END_VAR
VAR_OUTPUT
    nDays    : INT;   // 距重新标定的天数（负值 = 已超标）[天] / Days until recalibration, negative means overdue
    bOverdue : BOOL;  // 已超期 [-] / Recalibration overdue
END_VAR
VAR
    _fRate : REAL;  // 漂移速率绝对值 [单位/天] / Absolute drift rate
    _fEla  : REAL;  // 已标定天数 [天] / Days elapsed since the last calibration
    _fRem  : REAL;  // 允许剩余漂移 [单位] / Allowed remaining drift
    _fDay  : REAL;  // 剩余天数（钳定前）[天] / Remaining days before clamping
END_VAR
VAR CONSTANT
    DL_RDC_SEC_DAY  : REAL := 86400.0;   // 每天的秒数 [s/天] / Seconds per day
    DL_RDC_MS_S     : REAL := 1000.0;    // 毫秒 → 秒换算系数 [ms/s] / Milliseconds per second
    DL_RDC_RATE_EPS : REAL := 1.0E-9;    // 漂移速率判零下限 [单位/天] / Zero floor of the drift rate
    DL_RDC_DMAX     : REAL := 32000.0;   // 实数域钳制上限（INT 可表）[天] / Real domain clamp bound
    DL_RDC_SENTINEL : INT  := 32767;     // 永不超期哨兵值 [天] / Sentinel value for never overdue
END_VAR

(* 段 0：出口预置安全侧（0 天 = 立即需标定，N1/N3） *)
FC_DL_AnalyzerRecalDaysCalc := FALSE;
nDays := 0;  bOverdue := TRUE;

(* 段 1：非有限闸（三个浮点入参） *)
IF (fDriftRate <> fDriftRate) OR (fDriftLimit <> fDriftLimit) OR (fDriftNow <> fDriftNow) THEN RETURN; END_IF

(* 段 2：组态闸（允许漂移上限必须为正，否则按已超期） *)
IF fDriftLimit <= 0.0 THEN RETURN; END_IF

(* 段 3：漂移速率判零闸（近零速率 → 永不超期哨兵） *)
_fRate := ABS(fDriftRate);
IF _fRate <= DL_RDC_RATE_EPS THEN
    nDays := DL_RDC_SENTINEL;
    bOverdue := FALSE;                  // 漂移几乎为零：不报超期
    FC_DL_AnalyzerRecalDaysCalc := TRUE;
    RETURN;
END_IF

(* 段 4：剩余天数（除子已证 > 1E-9） *)
_fEla := TIME_TO_REAL(tSinceCal) / DL_RDC_MS_S / DL_RDC_SEC_DAY;
_fRem := fDriftLimit - ABS(fDriftNow);
_fDay := _fRem / _fRate - _fEla;
IF (_fDay <> _fDay) OR ((_fDay - _fDay) <> (_fDay - _fDay)) THEN RETURN; END_IF

(* 段 5：单一出口裁决（先钳后转型，判据与出口同源于 _fDay，N4/R23） *)
IF _fDay > DL_RDC_DMAX THEN
    _fDay := DL_RDC_DMAX;
ELSIF _fDay < (0.0 - DL_RDC_DMAX) THEN
    _fDay := 0.0 - DL_RDC_DMAX;         // 负向钳定：保留超期方向
END_IF
nDays := REAL_TO_INT(_fDay);
bOverdue := (_fDay < 0.0);
FC_DL_AnalyzerRecalDaysCalc := NOT bOverdue;
END_FUNCTION

(* ---- FC_DL_AsrsCycleTimeCalc.st ---- *)
(*
  DL Factory R83 | FC_DL_AsrsCycleTimeCalc
  功能：按梯形速度曲线分别算堆垛机行走与升降时间，取慢者加货叉时间得单循环。
  开源溯源：无（clean-room 自研，依据公开工艺公式，来源=行业通用公式，许可证=MIT，借鉴点=公式结构）
  规则：R1-R21 全遵守
*)
FUNCTION FC_DL_AsrsCycleTimeCalc : REAL
VAR_INPUT
    fTravelM   : REAL; // 巷道行走距离 [m] / Aisle travel distance [m]
    fTravelMps : REAL; // 行走最大速度 [m/s] / Travel maximum speed [m/s]
    fTravelAcc : REAL; // 行走加速度 [m/s²] / Travel acceleration [m/s^2]
    fLiftM     : REAL; // 升降行程 [m] / Lift stroke [m]
    fLiftMps   : REAL; // 升降最大速度 [m/s] / Lift maximum speed [m/s]
    fLiftAcc   : REAL; // 升降加速度 [m/s²] / Lift acceleration [m/s^2]
    fForkSec   : REAL; // 货叉单次伸缩时间 [s] / Fork stroke time [s]
END_VAR
VAR_OUTPUT
    fTravelS : REAL; // 行走段耗时 [s] / Travel leg time [s]
    fLiftS   : REAL; // 升降段耗时 [s] / Lift leg time [s]
    fCycleS  : REAL; // 单循环作业时间（两轴取大 + 货叉）[s] / Single cycle time [s]
    xValid   : BOOL; // 计算有效性标志 / Calculation validity flag
END_VAR
VAR
    fCritTravelM : REAL; // 行走达速临界距离 [m] / Travel distance to reach max speed [m]
    fCritLiftM   : REAL; // 升降达速临界距离 [m] / Lift distance to reach max speed [m]
END_VAR
fTravelS := 0.0; fLiftS := 0.0; fCycleS := 0.0; xValid := FALSE;  // 出口预置（R256）
// 非有限拦截 + 量纲自检 + 速度/加速度零闸（R4/R20/R21）
IF NOT (fTravelM > -1.0E30 AND fTravelM < 1.0E30) OR NOT (fTravelMps > -1.0E30 AND fTravelMps < 1.0E30) OR NOT (fTravelAcc > -1.0E30 AND fTravelAcc < 1.0E30) OR NOT (fLiftM > -1.0E30 AND fLiftM < 1.0E30) OR NOT (fLiftMps > -1.0E30 AND fLiftMps < 1.0E30) OR NOT (fLiftAcc > -1.0E30 AND fLiftAcc < 1.0E30) OR NOT (fForkSec > -1.0E30 AND fForkSec < 1.0E30) OR fTravelM < 0.0 OR fLiftM < 0.0 OR fForkSec < 0.0 OR fTravelMps <= 0.0 OR fLiftMps <= 0.0 OR fTravelAcc <= 0.0 OR fLiftAcc <= 0.0 THEN
    FC_DL_AsrsCycleTimeCalc := -1.0; RETURN;   // 哨兵 -1：非有限或量纲越界 / Sentinel -1
END_IF
// 行走段：临界距离 v²/a，超过则梯形曲线，否则三角曲线（t = 2√(d/a)）
fCritTravelM := (fTravelMps * fTravelMps) / fTravelAcc;   // 临界距离 [m] / Critical distance [m]
IF fTravelM >= fCritTravelM THEN
    fTravelS := fTravelM / fTravelMps + fTravelMps / fTravelAcc; // 梯形：d/v + v/a，量纲 s
ELSE
    fTravelS := 2.0 * SQRT(fTravelM / fTravelAcc);   // 三角：未达速，2√(d/a)，被除数已非负（R4）
END_IF
// 升降段：同一梯形/三角判据，参数完全独立
fCritLiftM := (fLiftMps * fLiftMps) / fLiftAcc;            // 临界距离 [m] / Critical distance [m]
IF fLiftM >= fCritLiftM THEN fLiftS := fLiftM / fLiftMps + fLiftMps / fLiftAcc; ELSE fLiftS := 2.0 * SQRT(fLiftM / fLiftAcc); END_IF  // 升降梯形/三角 [s]
// 单循环：两轴并行取较慢者，再串行加货叉伸缩（s + s = s）
IF fTravelS >= fLiftS THEN
    fCycleS := fTravelS + fForkSec; // 行走为瓶颈 [s] / Travel is the bottleneck
ELSE
    fCycleS := fLiftS + fForkSec;   // 升降为瓶颈 [s] / Lift is the bottleneck
END_IF
xValid := TRUE;                            // 链路有效 / Chain valid
FC_DL_AsrsCycleTimeCalc := fCycleS;        // 返回单循环时间 [s] / Return single cycle time [s]
END_FUNCTION

(* ---- FC_DL_BarrelRotationRpmCalc.st ---- *)
(*
  DL Factory R83 | FC_DL_BarrelRotationRpmCalc
  功能：按滚筒内径与零件贴壁尺寸算临界转速，并给出实际转速与临界转速之比。
  开源溯源：无（clean-room 自研，依据公开工艺公式，来源=行业通用公式，许可证=MIT，借鉴点=公式结构）
  规则：R1-R21 全遵守
*)
FUNCTION FC_DL_BarrelRotationRpmCalc : REAL
VAR_INPUT
    fBarrelDiaMm : REAL; // 滚筒内径 [mm] / Barrel inner diameter [mm]
    fRpm         : REAL; // 实测滚筒转速 [rpm] / Measured barrel speed [rpm]
    fPartDiaMm   : REAL; // 零件特征尺寸（贴壁层厚近似）[mm] / Part characteristic size [mm]
    fFillPct     : REAL; // 装载率（0~60）[%] / Barrel fill ratio [%]
END_VAR
VAR_OUTPUT
    fCritRpm  : REAL; // 临界转速（物料离心贴壁起始）[rpm] / Critical speed [rpm]
    fRpmRatio : REAL; // 转速比（实际÷临界，工艺宜 0.3~0.6）[-] / Speed ratio, window 0.3 to 0.6
    xValid    : BOOL; // 计算有效性标志 / Calculation validity flag
END_VAR
VAR
    fEffDiaM : REAL; // 有效内径（扣除贴壁层）[m] / Effective inner diameter [m]
    fSqrtD   : REAL; // 有效内径平方根 [m^0.5] / Square root of effective diameter [m^0.5]
END_VAR
fCritRpm := 0.0; fRpmRatio := 0.0; xValid := FALSE;  // 出口预置（R256）
// 非有限拦截 + 几何量纲自检（R20/R21）
IF NOT (fBarrelDiaMm > -1.0E30 AND fBarrelDiaMm < 1.0E30) OR NOT (fRpm > -1.0E30 AND fRpm < 1.0E30) OR NOT (fPartDiaMm > -1.0E30 AND fPartDiaMm < 1.0E30) OR NOT (fFillPct > -1.0E30 AND fFillPct < 1.0E30) OR fBarrelDiaMm <= 0.0 OR fRpm < 0.0 OR fPartDiaMm < 0.0 OR fPartDiaMm >= fBarrelDiaMm THEN
    FC_DL_BarrelRotationRpmCalc := -1.0; RETURN;  // 哨兵 -1：非有限或几何越界 / Sentinel -1
END_IF
// 装载率域闸：0~60% 之外钳位（超装将改变物料运动形态）
IF fFillPct < 0.0 THEN fFillPct := 0.0; ELSIF fFillPct > 60.0 THEN fFillPct := 60.0; END_IF
// 有效内径：滚筒内径扣减两层零件贴壁厚度，mm ÷ 1000 = m（量纲自洽）
fEffDiaM := (fBarrelDiaMm - 2.0 * fPartDiaMm) / 1000.0; // 有效内径 [m] / Effective inner diameter
// 开方前非负闸（R4），再按经验式 n_c = 42.3 / √D 算临界转速（D 单位 m，n_c 单位 rpm）
IF fEffDiaM > 0.0 THEN
    fSqrtD := SQRT(fEffDiaM);       // 内径平方根 [m^0.5] / Square root of diameter
    IF ABS(fSqrtD) > 1.0E-9 THEN fCritRpm := 42.3 / fSqrtD; ELSE fCritRpm := 0.0; END_IF
ELSE
    fCritRpm := 0.0;                // 内径非正不可算，缺省零 / Non-positive diameter, default zero
END_IF
// 转速比：实际 ÷ 临界，临界转速分母显式零闸（R4/R21）
IF ABS(fCritRpm) > 1.0E-9 THEN      // 临界转速分母显式零闸 / Explicit zero gate
    fRpmRatio := fRpm / fCritRpm;   // 转速比 [-]/ Speed ratio
ELSE
    fRpmRatio := 0.0;               // 除零防御缺省 / Divide-by-zero default
END_IF
xValid := TRUE; FC_DL_BarrelRotationRpmCalc := fRpmRatio;  // 返回转速比 [-] / Return speed ratio
END_FUNCTION
